// TIA Portal project "000_empty" (V21)

(* hardware
DEVICE "PLC_1"  S7-1500 station
   slot 0: "Rail_0"  Rack  6ES7 590-1***0-0AA0
   slot 1: "PLC_1"  CPU 1513-1 PN  6ES7 513-1AL02-0AB0  V2.9
      slot 3: "CPU display_1"  6ES7591-1AA00-0AA0
      slot 32768: "PROFINET interface_1"  X1
         slot 32769: "Port_1"  X1 P1
         slot 32770: "Port_2"  X1 P2
      slot 34817: "Virtual CP interface port_1"  Virtual CP interface port  Virtual CP interface port
DEVICE "HMI_TP900"  TP900 Comfort
   slot 0: "HMI_TP900"  TP900 Comfort  6AV2 124-0JC01-0AX0  17.0.0.0
   slot 1: "HMI_TP900"  TP900 Comfort  6AV2 124-0JC01-0AX0  17.0.0.0
   slot 5: "HMI_TP900.IE_CP_1"  PROFINET Interface  17.0.0.0
      slot 1: "PROFINET Interface_1"  PROFINET Interface
         slot 1: "Port_1"  Port
         slot 2: "Port_2"  Port
   slot 7: "HMI_TP900.MPI/DP_CP_1"  MPI/DP Interface  17.0.0.0
DEVICE "HMI_PCADV"  SIMATIC PC station
   slot 0: "SIMATIC PC station"  Rail  SIMATIC PC-Station  V1.0
      slot 125: "Stationmanager"  Station_Manager  V6.0.4
   slot 1: "HMI_RT_1"  WinCC RT Advanced  6AV2 104-0xxxx-xxxx  17.0.0.0
      slot 33792: "Computer interface"  Host interface
   slot 2: "IE_general_1"  IE General  IE_CP  V8.2.0
      slot 1: "PROFINET interface"  IEGeneral.Interface.8.2.0
DEVICE "HMI_TP900S"  TP900 Comfort
   slot 0: "HMI_TP900S"  TP900 Comfort  6AV2 124-0JC01-0AX0  17.0.0.0
   slot 1: "HMI_TP900S"  TP900 Comfort  6AV2 124-0JC01-0AX0  17.0.0.0
   slot 5: "HMI_TP900S.IE_CP_1"  PROFINET Interface  17.0.0.0
      slot 1: "PROFINET Interface_1"  PROFINET Interface
         slot 1: "Port_1"  Port
         slot 2: "Port_2"  Port
   slot 7: "HMI_TP900S.MPI/DP_CP_1"  MPI/DP Interface  17.0.0.0
DEVICE "HMI_TP1200"  TP1200 Comfort
   slot 0: "HMI_TP1200"  TP1200 Comfort  6AV2 124-0MC01-0AX0  17.0.0.0
   slot 1: "HMI_TP1200"  TP1200 Comfort  6AV2 124-0MC01-0AX0  17.0.0.0
   slot 5: "HMI_TP1200.IE_CP_1"  PROFINET Interface  17.0.0.0
      slot 1: "PROFINET Interface_1"  PROFINET Interface
         slot 1: "Port_1"  Port
         slot 2: "Port_2"  Port
   slot 7: "HMI_TP1200.MPI/DP_CP_1"  MPI/DP Interface  17.0.0.0
*)

// ===== PLC "PLC_1"  CPU 1513-1 PN =====

VAR_GLOBAL   // PLC tag table "Default tag table"
   "Plc_Bool" AT %M100.0 : Bool;
   "Plc_Int" AT %MW102 : Int;
   "Plc_Real" AT %MD104 : Real;
   "Plc_Byte" AT %MB108 : Byte;
END_VAR

ORGANIZATION_BLOCK "Main"   // OB1, LAD, ProgramCycle
TITLE = "Main Program Sweep (Cycle)"
{ S7_Optimized_Access := 'TRUE' }
VERSION : 0.1
   VAR_INPUT
      Initial_Call : Bool;   // Initial call of this OB
      Remanence : Bool;   // =True, if remanent data are available
   END_VAR
BEGIN
END_ORGANIZATION_BLOCK

(* ===== HMI "HMI_TP900" =====
system functions are stored by id; their names below are inferred from use
connection "HMI_Connection_1": ETHERNET, S7_1500_OMS

HMI tags "Default tag table"
   "Hmi_Bool" : Bool, internal
   "Hmi_Int" : Int, internal
   "Hmi_Real" : Real, internal
   "Hmi_String" : WString[254], internal
   "Ext_Bool" : Bool = PLC Plc_Bool AT %M100.0, 1 s
   "Ext_Int" : Int = PLC Plc_Int AT %MW102, 1 s
   "Ext_Real" : Real = PLC Plc_Real AT %MD104, 1 s
   "Ext_Byte" : Byte = PLC Plc_Byte AT %MB108, 1 s

HMI tags "C03_Tags"
   "D_State" : Int, internal
   "D_Bool" : Bool, internal
   "D_SInt" : SInt, internal
   "D_Int" : Int, internal
   "D_DInt" : DInt, internal
   "D_USInt" : USInt, internal
   "D_UInt" : UInt, internal
   "D_UDInt" : UDInt, internal
   "D_Real" : Real, internal
   "D_LReal" : LReal, internal
   "D_String" : WString[254], internal
   "D_DateTime" : DateTime, internal
   "D_Pct" : Int, internal
   "D_Range" : Int, internal
   "D_Bits" : Int, internal
   "D_Vis" : Bool, internal
   "D_En" : Bool, internal
   "D_X" : Int, internal
   "D_Y" : Int, internal
   "D_Max" : Real, internal
   "D_Min" : Real, internal
   "D_TL" : Int, internal
   "D_BarR" : Real, internal

text list "TL_Value": -100..-1 'Negative (-100..-1)'; 0 'Zero'; 1..9 'One to nine'; 10 'Ten: Ünïcödé äöüß ÄÖÜ €'; 32000 'Undefined value (default entry)'

text list "TL_Bit": 0 'Off (0)'; 1 'On (1)'

text list "TL_BitNo": 0 'Bit 0 set'; 1 'Bit 1 set'; 2 'Bit 2 set'; 3 'Bit 3 set'

graphic list "GL_Bit": 0 'G_EMF'; 1 'G_WMF'

graphic list "GL_BitNo": 0 'G_PNG'; 1 'G_JPG'; 2 'G_BMP'; 3 'G_TIF'

graphic list "GL_Value": -100..-1 'G_GIF'; 0 'G_PNG'; 1..9 'G_JPG'; 10 'G_BMP'; 32000 'G_SVG'

SlideinScreen "GraphX_Slidein_Top" 800x120
   TextField "SI_Title" at 10,10 size 300x20; Text 'Slide-in screen Top'
   Bar "SI_Bar" at 330,10 size 200x40
      ProcessValue <- "D_Pct"
   IOField "SI_Value" at 560,10 size 120x30; FormatPattern s99999
      ProcessValue <- "D_Int"

screen "All_Objects" 800x480
   TextField "TextField_1" at 680,10 size 100x30; Text 'Text'
   GraphicView "GraphicView_1" at 10,80 size 100x60
   IOField "IOField_1" at 130,80 size 100x30
   Button "Button_1" at 250,80 size 100x40; TextOff 'Text'
   SymbolicIOField "SymbolicIOField_1" at 370,80 size 120x30; TextOff '0'; TextOn '1'
   GraphicIOField "GraphicIOField_1" at 510,80 size 60x60
   DateTimeField "DateTimeField_1" at 590,80 size 160x30
   Bar "Bar_1" at 10,160 size 40x120
   Switch "Switch_1" at 70,160 size 120x40; CaptionText 'Switch'; TextOff '0'; TextOn '1'
   SymbolLibrary "SymbolLibrary_1" at 210,160 size 60x60
   Slider "Slider_1" at 290,160 size 60x160; Caption 'SIMATIC'
   Gauge "Gauge_1" at 370,160 size 150x150; CaptionText 'SIMATIC'
   Clock "Clock_1" at 540,160 size 150x150

screen "Ctl_01_AlarmView" 800x480, template "Nav"
   AlarmView "Alarm view_1" at 3,3 size 600x300

screen "Ctl_02_TrendView" 800x480, template "Nav"
   TrendView "Trend view_1" at 3,3 size 600x300

screen "Ctl_03_UserView" 800x480, template "Nav"
   UserView "User view_1" at 3,3 size 480x240

screen "Ctl_04_HtmlBrowser" 800x480, template "Nav"
   HTMLBrowser "HTML browser_1" at 3,3 size 192x192

screen "Ctl_05_WatchTable" 800x480, template "Nav"
   StatusForce "Watch table_1" at 3,3 size 600x300; ToolTipText 'Text'

screen "Ctl_06_SmartClientView" 800x480, template "Nav"
   SmartClientView "Sm@rtClient view_1" at 3,3 size 320x240

screen "Ctl_07_RecipeView" 800x480, template "Nav"
   RecipeView "Recipe view_1" at 3,3 size 400x330

screen "Ctl_09_SysDiagView" 800x480, template "Nav"
   SysDiagControl "System diagnostics view_1" at 3,3 size 600x300

screen "Ctl_10_MediaPlayer" 800x480, template "Nav"
   MediaPlayer "Media Player_1" at 3,3 size 240x240

screen "Ctl_15_CameraView" 800x480, template "Nav"
   CameraControl "Camera view_1" at 3,3 size 320x240

screen "Ctl_16_PdfView" 800x480, template "Nav"
   PDFView "PDFView_1" at 3,3 size 320x240

Template "Nav" 800x480
   Button "Nav_01" at 770,2 size 28x22; TextOff 'Text'
      on Click: ActivateScreen("Ctl_01_AlarmView", 0)
   Button "Nav_02" at 770,28 size 28x22; TextOff 'Text'
      on Click: ActivateScreen("Ctl_02_TrendView", 0)
   Button "Nav_03" at 770,54 size 28x22; TextOff 'Text'
      on Click: ActivateScreen("Ctl_03_UserView", 0)
   Button "Nav_04" at 770,80 size 28x22; TextOff 'Text'
      on Click: ActivateScreen("Ctl_04_HtmlBrowser", 0)
   Button "Nav_05" at 770,106 size 28x22; TextOff 'Text'
      on Click: ActivateScreen("Ctl_05_WatchTable", 0)
   Button "Nav_06" at 770,132 size 28x22; TextOff 'Text'
      on Click: ActivateScreen("Ctl_06_SmartClientView", 0)
   Button "Nav_07" at 770,158 size 28x22; TextOff 'Text'
      on Click: ActivateScreen("Ctl_07_RecipeView", 0)
   Button "Nav_09" at 770,210 size 28x22; TextOff 'Text'
      on Click: ActivateScreen("Ctl_09_SysDiagView", 0)
   Button "Nav_10" at 770,236 size 28x22; TextOff 'Text'
      on Click: ActivateScreen("Ctl_10_MediaPlayer", 0)
   Button "Nav_15" at 770,366 size 28x22; TextOff 'Text'
      on Click: ActivateScreen("Ctl_15_CameraView", 0)
   Button "Nav_16" at 770,392 size 28x22; TextOff 'Text'
      on Click: ActivateScreen("Ctl_16_PdfView", 0)
   Button "Nav_17" at 770,418 size 28x22; TextOff 'Text'
      on Click: ActivateScreen("All_Objects", 0)

screen "P_Line_1" 800x480
   TextField "Label_Default" at 10,62 size 108x16; Text 'Default'
   TextField "Label_BackColor" at 120,62 size 108x16; Text 'BackColor'
   TextField "Label_Color" at 230,62 size 108x16; Text 'Color'
   TextField "Label_EndStyle" at 340,62 size 108x16; Text 'EndStyle'
   TextField "Label_EndStyle_2" at 450,62 size 108x16; Text 'EndStyle_2'
   TextField "Label_EndStyle_3" at 560,62 size 108x16; Text 'EndStyle_3'
   TextField "Label_EndStyle_4" at 670,62 size 108x16; Text 'EndStyle_4'
   TextField "Label_EndStyle_5" at 10,138 size 108x16; Text 'EndStyle_5'
   TextField "Label_FillStyle" at 120,138 size 108x16; Text 'FillStyle'
   TextField "Label_Flashing" at 230,138 size 108x16; Text 'Flashing'
   TextField "Label_LineEndShapeStyle_2" at 340,138 size 108x16; Text 'LineEndShapeStyle_2'
   TextField "Label_LineWidth" at 450,138 size 108x16; Text 'LineWidth'
   TextField "Label_StartStyle" at 560,138 size 108x16; Text 'StartStyle'
   TextField "Label_StartStyle_2" at 670,138 size 108x16; Text 'StartStyle_2'
   TextField "Label_StartStyle_3" at 10,214 size 108x16; Text 'StartStyle_3'
   TextField "Label_StartStyle_4" at 120,214 size 108x16; Text 'StartStyle_4'
   TextField "Label_StartStyle_5" at 230,214 size 108x16; Text 'StartStyle_5'
   TextField "Label_Style" at 340,214 size 108x16; Text 'Style'
   TextField "Label_Style_2" at 450,214 size 108x16; Text 'Style_2'
   TextField "Label_Style_3" at 560,214 size 108x16; Text 'Style_3'
   TextField "Label_Style_4" at 670,214 size 108x16; Text 'Style_4'
   TextField "Label_UseDesignColorSchema" at 10,290 size 108x16; Text 'UseDesignColorSchema'
   Button "Next" at 758,456 size 40x22; TextOff 'Text'
      on Click: ActivateScreen("P_Polyline_1", 0)

screen "P_Polyline_1" 800x480
   TextField "Label_Default" at 10,62 size 108x16; Text 'Default'
   TextField "Label_BackColor" at 120,62 size 108x16; Text 'BackColor'
   TextField "Label_Color" at 230,62 size 108x16; Text 'Color'
   TextField "Label_EndStyle" at 340,62 size 108x16; Text 'EndStyle'
   TextField "Label_EndStyle_2" at 450,62 size 108x16; Text 'EndStyle_2'
   TextField "Label_EndStyle_3" at 560,62 size 108x16; Text 'EndStyle_3'
   TextField "Label_EndStyle_4" at 670,62 size 108x16; Text 'EndStyle_4'
   TextField "Label_EndStyle_5" at 10,138 size 108x16; Text 'EndStyle_5'
   TextField "Label_FillStyle" at 120,138 size 108x16; Text 'FillStyle'
   TextField "Label_Flashing" at 230,138 size 108x16; Text 'Flashing'
   TextField "Label_LineEndShapeStyle_2" at 340,138 size 108x16; Text 'LineEndShapeStyle_2'
   TextField "Label_LineWidth" at 450,138 size 108x16; Text 'LineWidth'
   TextField "Label_StartStyle" at 560,138 size 108x16; Text 'StartStyle'
   TextField "Label_StartStyle_2" at 670,138 size 108x16; Text 'StartStyle_2'
   TextField "Label_StartStyle_3" at 10,214 size 108x16; Text 'StartStyle_3'
   TextField "Label_StartStyle_4" at 120,214 size 108x16; Text 'StartStyle_4'
   TextField "Label_StartStyle_5" at 230,214 size 108x16; Text 'StartStyle_5'
   TextField "Label_Style" at 340,214 size 108x16; Text 'Style'
   TextField "Label_Style_2" at 450,214 size 108x16; Text 'Style_2'
   TextField "Label_Style_3" at 560,214 size 108x16; Text 'Style_3'
   TextField "Label_Style_4" at 670,214 size 108x16; Text 'Style_4'
   TextField "Label_UseDesignColorSchema" at 10,290 size 108x16; Text 'UseDesignColorSchema'
   Button "Next" at 758,456 size 40x22; TextOff 'Text'
      on Click: ActivateScreen("P_Polygon_1", 0)

screen "P_Polygon_1" 800x480
   TextField "Label_Default" at 10,62 size 108x16; Text 'Default'
   TextField "Label_BackColor" at 120,62 size 108x16; Text 'BackColor'
   TextField "Label_BackFillStyle" at 230,62 size 108x16; Text 'BackFillStyle'
   TextField "Label_BorderColor" at 340,62 size 108x16; Text 'BorderColor'
   TextField "Label_BorderWidth" at 450,62 size 108x16; Text 'BorderWidth'
   TextField "Label_EdgeStyle" at 560,62 size 108x16; Text 'EdgeStyle'
   TextField "Label_EdgeStyle_2" at 670,62 size 108x16; Text 'EdgeStyle_2'
   TextField "Label_EdgeStyle_3" at 10,138 size 108x16; Text 'EdgeStyle_3'
   TextField "Label_EdgeStyle_4" at 120,138 size 108x16; Text 'EdgeStyle_4'
   TextField "Label_Flashing" at 230,138 size 108x16; Text 'Flashing'
   TextField "Label_UseDesignColorSchema" at 340,138 size 108x16; Text 'UseDesignColorSchema'
   Button "Next" at 758,456 size 40x22; TextOff 'Text'
      on Click: ActivateScreen("P_Ellipse_1", 0)

screen "P_Ellipse_1" 800x480
   TextField "Label_Default" at 10,62 size 108x16; Text 'Default'
   TextField "Label_BackColor" at 120,62 size 108x16; Text 'BackColor'
   TextField "Label_BackFillStyle" at 230,62 size 108x16; Text 'BackFillStyle'
   TextField "Label_BorderColor" at 340,62 size 108x16; Text 'BorderColor'
   TextField "Label_BorderWidth" at 450,62 size 108x16; Text 'BorderWidth'
   TextField "Label_EdgeStyle" at 560,62 size 108x16; Text 'EdgeStyle'
   TextField "Label_EdgeStyle_2" at 670,62 size 108x16; Text 'EdgeStyle_2'
   TextField "Label_EdgeStyle_3" at 10,138 size 108x16; Text 'EdgeStyle_3'
   TextField "Label_EdgeStyle_4" at 120,138 size 108x16; Text 'EdgeStyle_4'
   TextField "Label_Flashing" at 230,138 size 108x16; Text 'Flashing'
   TextField "Label_UseDesignColorSchema" at 340,138 size 108x16; Text 'UseDesignColorSchema'
   Button "Next" at 758,456 size 40x22; TextOff 'Text'
      on Click: ActivateScreen("P_Circle_1", 0)

screen "P_Circle_1" 800x480
   TextField "Label_Default" at 10,62 size 58x16; Text 'Default'
   TextField "Label_BackColor" at 70,62 size 58x16; Text 'BackColor'
   TextField "Label_BackFillStyle" at 130,62 size 58x16; Text 'BackFillStyle'
   TextField "Label_BorderColor" at 190,62 size 58x16; Text 'BorderColor'
   TextField "Label_BorderWidth" at 250,62 size 58x16; Text 'BorderWidth'
   TextField "Label_EdgeStyle" at 310,62 size 58x16; Text 'EdgeStyle'
   TextField "Label_EdgeStyle_2" at 370,62 size 58x16; Text 'EdgeStyle_2'
   TextField "Label_EdgeStyle_3" at 430,62 size 58x16; Text 'EdgeStyle_3'
   TextField "Label_EdgeStyle_4" at 490,62 size 58x16; Text 'EdgeStyle_4'
   TextField "Label_Flashing" at 550,62 size 58x16; Text 'Flashing'
   TextField "Label_UseDesignColorSchema" at 610,62 size 58x16; Text 'UseDesignColorSchema'
   Button "Next" at 758,456 size 40x22; TextOff 'Text'
      on Click: ActivateScreen("P_Rectangle_1", 0)

screen "P_Rectangle_1" 800x480
   TextField "Label_Default" at 10,62 size 108x16; Text 'Default'
   TextField "Label_BackColor" at 120,62 size 108x16; Text 'BackColor'
   TextField "Label_BackFillStyle" at 230,62 size 108x16; Text 'BackFillStyle'
   TextField "Label_BorderColor" at 340,62 size 108x16; Text 'BorderColor'
   TextField "Label_BorderWidth" at 450,62 size 108x16; Text 'BorderWidth'
   TextField "Label_EdgeStyle" at 560,62 size 108x16; Text 'EdgeStyle'
   TextField "Label_EdgeStyle_2" at 670,62 size 108x16; Text 'EdgeStyle_2'
   TextField "Label_EdgeStyle_3" at 10,138 size 108x16; Text 'EdgeStyle_3'
   TextField "Label_EdgeStyle_4" at 120,138 size 108x16; Text 'EdgeStyle_4'
   TextField "Label_Flashing" at 230,138 size 108x16; Text 'Flashing'
   TextField "Label_RoundCornerHeight" at 340,138 size 108x16; Text 'RoundCornerHeight'
   TextField "Label_RoundCornerWidth" at 450,138 size 108x16; Text 'RoundCornerWidth'
   TextField "Label_UseDesignColorSchema" at 560,138 size 108x16; Text 'UseDesignColorSchema'
   Button "Next" at 758,456 size 40x22; TextOff 'Text'
      on Click: ActivateScreen("P_TextField_1", 0)

screen "P_TextField_1" 800x480
   TextField "Default" at 10,10 size 100x30; Text 'Text'
   TextField "Label_Default" at 10,42 size 108x16; Text 'Default'
   TextField "BackColor" at 120,10 size 100x30; Text 'Text'
   TextField "Label_BackColor" at 120,42 size 108x16; Text 'BackColor'
   TextField "BackFillStyle" at 230,10 size 100x30; Text 'Text'
   TextField "Label_BackFillStyle" at 230,42 size 108x16; Text 'BackFillStyle'
   TextField "BorderBackColor" at 340,10 size 100x30; Text 'Text'
   TextField "Label_BorderBackColor" at 340,42 size 108x16; Text 'BorderBackColor'
   TextField "BorderColor" at 450,10 size 100x30; Text 'Text'
   TextField "Label_BorderColor" at 450,42 size 108x16; Text 'BorderColor'
   TextField "BorderWidth" at 560,10 size 100x30; Text 'Text'
   TextField "Label_BorderWidth" at 560,42 size 108x16; Text 'BorderWidth'
   TextField "BottomMargin" at 670,10 size 100x30; Text 'Text'
   TextField "Label_BottomMargin" at 670,42 size 108x16; Text 'BottomMargin'
   TextField "CornerRadius" at 10,66 size 100x30; Text 'Text'
   TextField "Label_CornerRadius" at 10,98 size 108x16; Text 'CornerRadius'
   TextField "EdgeStyle" at 120,66 size 100x30; Text 'Text'
   TextField "Label_EdgeStyle" at 120,98 size 108x16; Text 'EdgeStyle'
   TextField "EdgeStyle_2" at 230,66 size 100x30; Text 'Text'
   TextField "Label_EdgeStyle_2" at 230,98 size 108x16; Text 'EdgeStyle_2'
   TextField "EdgeStyle_3" at 340,66 size 100x30; Text 'Text'
   TextField "Label_EdgeStyle_3" at 340,98 size 108x16; Text 'EdgeStyle_3'
   TextField "EdgeStyle_4" at 450,66 size 100x30; Text 'Text'
   TextField "Label_EdgeStyle_4" at 450,98 size 108x16; Text 'EdgeStyle_4'
   TextField "FitToLargest" at 560,66 size 100x30; Text 'Text'
   TextField "Label_FitToLargest" at 560,98 size 108x16; Text 'FitToLargest'
   TextField "Flashing" at 670,66 size 100x30; Text 'Text'
   TextField "Label_Flashing" at 670,98 size 108x16; Text 'Flashing'
   TextField "ForeColor" at 10,122 size 100x30; Text 'Text'
   TextField "Label_ForeColor" at 10,154 size 108x16; Text 'ForeColor'
   TextField "HorizontalAlignment" at 120,122 size 100x30; Text 'Text'
   TextField "Label_HorizontalAlignment" at 120,154 size 108x16; Text 'HorizontalAlignment'
   TextField "HorizontalAlignment_2" at 230,122 size 100x30; Text 'Text'
   TextField "Label_HorizontalAlignment_2" at 230,154 size 108x16; Text 'HorizontalAlignment_2'
   TextField "LeftMargin" at 340,122 size 100x30; Text 'Text'
   TextField "Label_LeftMargin" at 340,154 size 108x16; Text 'LeftMargin'
   TextField "RightMargin" at 450,122 size 100x30; Text 'Text'
   TextField "Label_RightMargin" at 450,154 size 108x16; Text 'RightMargin'
   TextField "TopMargin" at 560,122 size 100x30; Text 'Text'
   TextField "Label_TopMargin" at 560,154 size 108x16; Text 'TopMargin'
   TextField "UseDesignColorSchema" at 670,122 size 100x30; Text 'Text'
   TextField "Label_UseDesignColorSchema" at 670,154 size 108x16; Text 'UseDesignColorSchema'
   TextField "VerticalAlignment" at 10,178 size 100x30; Text 'Text'
   TextField "Label_VerticalAlignment" at 10,210 size 108x16; Text 'VerticalAlignment'
   TextField "VerticalAlignment_2" at 120,178 size 100x30; Text 'Text'
   TextField "Label_VerticalAlignment_2" at 120,210 size 108x16; Text 'VerticalAlignment_2'
   Button "Next" at 758,456 size 40x22; TextOff 'Text'
      on Click: ActivateScreen("P_GraphicView_1", 0)

screen "P_GraphicView_1" 800x480
   GraphicView "Default" at 10,10 size 100x60
   TextField "Label_Default" at 10,72 size 108x16; Text 'Default'
   GraphicView "BackColor" at 120,10 size 100x60
   TextField "Label_BackColor" at 120,72 size 108x16; Text 'BackColor'
   GraphicView "BackFillStyle" at 230,10 size 100x60
   TextField "Label_BackFillStyle" at 230,72 size 108x16; Text 'BackFillStyle'
   GraphicView "BorderColor" at 340,10 size 100x60
   TextField "Label_BorderColor" at 340,72 size 108x16; Text 'BorderColor'
   GraphicView "BorderWidth" at 450,10 size 100x60
   TextField "Label_BorderWidth" at 450,72 size 108x16; Text 'BorderWidth'
   GraphicView "EdgeStyle" at 560,10 size 100x60
   TextField "Label_EdgeStyle" at 560,72 size 108x16; Text 'EdgeStyle'
   GraphicView "EdgeStyle_2" at 670,10 size 100x60
   TextField "Label_EdgeStyle_2" at 670,72 size 108x16; Text 'EdgeStyle_2'
   GraphicView "EdgeStyle_3" at 10,96 size 100x60
   TextField "Label_EdgeStyle_3" at 10,158 size 108x16; Text 'EdgeStyle_3'
   GraphicView "EdgeStyle_4" at 120,96 size 100x60
   TextField "Label_EdgeStyle_4" at 120,158 size 108x16; Text 'EdgeStyle_4'
   GraphicView "FitToLargest" at 230,96 size 100x60
   TextField "Label_FitToLargest" at 230,158 size 108x16; Text 'FitToLargest'
   GraphicView "Flashing" at 340,96 size 100x60
   TextField "Label_Flashing" at 340,158 size 108x16; Text 'Flashing'
   GraphicView "TransparentColor" at 450,96 size 100x60
   TextField "Label_TransparentColor" at 450,158 size 108x16; Text 'TransparentColor'
   GraphicView "UseTransparentColor" at 560,96 size 100x60
   TextField "Label_UseTransparentColor" at 560,158 size 108x16; Text 'UseTransparentColor'
   Button "Next" at 758,456 size 40x22; TextOff 'Text'
      on Click: ActivateScreen("P_IOField_1", 0)

screen "P_Button_1" 800x480
   Button "Default" at 10,10 size 100x40; TextOff 'Text'
   TextField "Label_Default" at 10,52 size 108x16; Text 'Default'
   Button "BackColor" at 120,10 size 100x40; TextOff 'Text'
   TextField "Label_BackColor" at 120,52 size 108x16; Text 'BackColor'
   Button "BackFillStyle" at 230,10 size 100x40; TextOff 'Text'
   TextField "Label_BackFillStyle" at 230,52 size 108x16; Text 'BackFillStyle'
   Button "BorderBackColor" at 340,10 size 100x40; TextOff 'Text'
   TextField "Label_BorderBackColor" at 340,52 size 108x16; Text 'BorderBackColor'
   Button "BorderColor" at 450,10 size 100x40; TextOff 'Text'
   TextField "Label_BorderColor" at 450,52 size 108x16; Text 'BorderColor'
   Button "BorderWidth" at 560,10 size 100x40; TextOff 'Text'
   TextField "Label_BorderWidth" at 560,52 size 108x16; Text 'BorderWidth'
   Button "CornerRadius" at 670,10 size 100x40; TextOff 'Text'
   TextField "Label_CornerRadius" at 670,52 size 108x16; Text 'CornerRadius'
   Button "EdgeStyle" at 10,76 size 100x40; TextOff 'Text'
   TextField "Label_EdgeStyle" at 10,118 size 108x16; Text 'EdgeStyle'
   Button "EdgeStyle_2" at 120,76 size 100x40; TextOff 'Text'
   TextField "Label_EdgeStyle_2" at 120,118 size 108x16; Text 'EdgeStyle_2'
   Button "EdgeStyle_3" at 230,76 size 100x40; TextOff 'Text'
   TextField "Label_EdgeStyle_3" at 230,118 size 108x16; Text 'EdgeStyle_3'
   Button "EdgeStyle_4" at 340,76 size 100x40; TextOff 'Text'
   TextField "Label_EdgeStyle_4" at 340,118 size 108x16; Text 'EdgeStyle_4'
   Button "FirstGradientColor" at 450,76 size 100x40; TextOff 'Text'
   TextField "Label_FirstGradientColor" at 450,118 size 108x16; Text 'FirstGradientColor'
   Button "FirstGradientOffset" at 560,76 size 100x40; TextOff 'Text'
   TextField "Label_FirstGradientOffset" at 560,118 size 108x16; Text 'FirstGradientOffset'
   Button "FitToLargest" at 670,76 size 100x40; TextOff 'Text'
   TextField "Label_FitToLargest" at 670,118 size 108x16; Text 'FitToLargest'
   Button "Flashing" at 10,142 size 100x40; TextOff 'Text'
   TextField "Label_Flashing" at 10,184 size 108x16; Text 'Flashing'
   Button "FocusColor" at 120,142 size 100x40; TextOff 'Text'
   TextField "Label_FocusColor" at 120,184 size 108x16; Text 'FocusColor'
   Button "FocusWidth" at 230,142 size 100x40; TextOff 'Text'
   TextField "Label_FocusWidth" at 230,184 size 108x16; Text 'FocusWidth'
   Button "ForeColor" at 340,142 size 100x40; TextOff 'Text'
   TextField "Label_ForeColor" at 340,184 size 108x16; Text 'ForeColor'
   Button "HorizontalAlignment" at 450,142 size 100x40; TextOff 'Text'
   TextField "Label_HorizontalAlignment" at 450,184 size 108x16; Text 'HorizontalAlignment'
   Button "HorizontalAlignment_2" at 560,142 size 100x40; TextOff 'Text'
   TextField "Label_HorizontalAlignment_2" at 560,184 size 108x16; Text 'HorizontalAlignment_2'
   Button "HorizontalPictureAlignment" at 670,142 size 100x40; TextOff 'Text'
   TextField "Label_HorizontalPictureAlignment" at 670,184 size 108x16; Text 'HorizontalPictureAlignment'
   Button "HorizontalPictureAlignment_2" at 10,208 size 100x40; TextOff 'Text'
   TextField "Label_HorizontalPictureAlignment_2" at 10,250 size 108x16; Text 'HorizontalPictureAlignment_2'
   Button "MiddleGradientColor" at 120,208 size 100x40; TextOff 'Text'
   TextField "Label_MiddleGradientColor" at 120,250 size 108x16; Text 'MiddleGradientColor'
   Button "Mode_5" at 230,208 size 100x40; TextOff 'Text'
   TextField "Label_Mode_5" at 230,250 size 108x16; Text 'Mode_5'
   Button "Mode_7" at 340,208 size 100x40; TextOff 'Text'
   TextField "Label_Mode_7" at 340,250 size 108x16; Text 'Mode_7'
   Button "PictureAreaBottomMargin" at 450,208 size 100x40; TextOff 'Text'
   TextField "Label_PictureAreaBottomMargin" at 450,250 size 108x16; Text 'PictureAreaBottomMargin'
   Button "PictureAreaLeftMargin" at 560,208 size 100x40; TextOff 'Text'
   TextField "Label_PictureAreaLeftMargin" at 560,250 size 108x16; Text 'PictureAreaLeftMargin'
   Button "PictureAreaRightMargin" at 670,208 size 100x40; TextOff 'Text'
   TextField "Label_PictureAreaRightMargin" at 670,250 size 108x16; Text 'PictureAreaRightMargin'
   Button "PictureAreaTopMargin" at 10,274 size 100x40; TextOff 'Text'
   TextField "Label_PictureAreaTopMargin" at 10,316 size 108x16; Text 'PictureAreaTopMargin'
   Button "SecondGradientColor" at 120,274 size 100x40; TextOff 'Text'
   TextField "Label_SecondGradientColor" at 120,316 size 108x16; Text 'SecondGradientColor'
   Button "SecondGradientOffset" at 230,274 size 100x40; TextOff 'Text'
   TextField "Label_SecondGradientOffset" at 230,316 size 108x16; Text 'SecondGradientOffset'
   Button "TextAreaBottomMargin" at 340,274 size 100x40; TextOff 'Text'
   TextField "Label_TextAreaBottomMargin" at 340,316 size 108x16; Text 'TextAreaBottomMargin'
   Button "TextAreaLeftMargin" at 450,274 size 100x40; TextOff 'Text'
   TextField "Label_TextAreaLeftMargin" at 450,316 size 108x16; Text 'TextAreaLeftMargin'
   Button "TextAreaRightMargin" at 560,274 size 100x40; TextOff 'Text'
   TextField "Label_TextAreaRightMargin" at 560,316 size 108x16; Text 'TextAreaRightMargin'
   Button "TextAreaTopMargin" at 670,274 size 100x40; TextOff 'Text'
   TextField "Label_TextAreaTopMargin" at 670,316 size 108x16; Text 'TextAreaTopMargin'
   Button "UseDesignColorSchema" at 10,340 size 100x40; TextOff 'Text'
   TextField "Label_UseDesignColorSchema" at 10,382 size 108x16; Text 'UseDesignColorSchema'
   Button "UseFirstGradient" at 120,340 size 100x40; TextOff 'Text'
   TextField "Label_UseFirstGradient" at 120,382 size 108x16; Text 'UseFirstGradient'
   Button "UseSecondGradient" at 230,340 size 100x40; TextOff 'Text'
   TextField "Label_UseSecondGradient" at 230,382 size 108x16; Text 'UseSecondGradient'
   Button "VerticalAlignment" at 340,340 size 100x40; TextOff 'Text'
   TextField "Label_VerticalAlignment" at 340,382 size 108x16; Text 'VerticalAlignment'
   Button "VerticalAlignment_2" at 450,340 size 100x40; TextOff 'Text'
   TextField "Label_VerticalAlignment_2" at 450,382 size 108x16; Text 'VerticalAlignment_2'
   Button "VerticalPictureAlignment" at 560,340 size 100x40; TextOff 'Text'
   TextField "Label_VerticalPictureAlignment" at 560,382 size 108x16; Text 'VerticalPictureAlignment'
   Button "VerticalPictureAlignment_2" at 670,340 size 100x40; TextOff 'Text'
   TextField "Label_VerticalPictureAlignment_2" at 670,382 size 108x16; Text 'VerticalPictureAlignment_2'
   Button "Next" at 758,456 size 40x22; TextOff 'Text'
      on Click: ActivateScreen("P_SymbolicIOField_1", 0)

screen "P_SymbolicIOField_1" 800x480
   SymbolicIOField "Default" at 10,10 size 120x30; TextOff '0'; TextOn '1'
   TextField "Label_Default" at 10,42 size 128x16; Text 'Default'
   SymbolicIOField "AboveUpperLimitColor" at 140,10 size 120x30; TextOff '0'; TextOn '1'
   TextField "Label_AboveUpperLimitColor" at 140,42 size 128x16; Text 'AboveUpperLimitColor'
   SymbolicIOField "BackColor" at 270,10 size 120x30; TextOff '0'; TextOn '1'
   TextField "Label_BackColor" at 270,42 size 128x16; Text 'BackColor'
   SymbolicIOField "BackFillStyle" at 400,10 size 120x30; TextOff '0'; TextOn '1'
   TextField "Label_BackFillStyle" at 400,42 size 128x16; Text 'BackFillStyle'
   SymbolicIOField "BelowLowerLimitColor" at 530,10 size 120x30; TextOff '0'; TextOn '1'
   TextField "Label_BelowLowerLimitColor" at 530,42 size 128x16; Text 'BelowLowerLimitColor'
   SymbolicIOField "BorderBackColor" at 660,10 size 120x30; TextOff '0'; TextOn '1'
   TextField "Label_BorderBackColor" at 660,42 size 128x16; Text 'BorderBackColor'
   SymbolicIOField "BorderColor" at 10,66 size 120x30; TextOff '0'; TextOn '1'
   TextField "Label_BorderColor" at 10,98 size 128x16; Text 'BorderColor'
   SymbolicIOField "BorderWidth" at 140,66 size 120x30; TextOff '0'; TextOn '1'
   TextField "Label_BorderWidth" at 140,98 size 128x16; Text 'BorderWidth'
   SymbolicIOField "BottomMargin" at 270,66 size 120x30; TextOff '0'; TextOn '1'
   TextField "Label_BottomMargin" at 270,98 size 128x16; Text 'BottomMargin'
   SymbolicIOField "CornerRadius" at 400,66 size 120x30; TextOff '0'; TextOn '1'
   TextField "Label_CornerRadius" at 400,98 size 128x16; Text 'CornerRadius'
   SymbolicIOField "CountVisibleItems" at 530,66 size 120x30; TextOff '0'; TextOn '1'
   TextField "Label_CountVisibleItems" at 530,98 size 128x16; Text 'CountVisibleItems'
   SymbolicIOField "EdgeStyle" at 660,66 size 120x30; TextOff '0'; TextOn '1'
   TextField "Label_EdgeStyle" at 660,98 size 128x16; Text 'EdgeStyle'
   SymbolicIOField "EdgeStyle_2" at 10,122 size 120x30; TextOff '0'; TextOn '1'
   TextField "Label_EdgeStyle_2" at 10,154 size 128x16; Text 'EdgeStyle_2'
   SymbolicIOField "EdgeStyle_3" at 140,122 size 120x30; TextOff '0'; TextOn '1'
   TextField "Label_EdgeStyle_3" at 140,154 size 128x16; Text 'EdgeStyle_3'
   SymbolicIOField "EdgeStyle_4" at 270,122 size 120x30; TextOff '0'; TextOn '1'
   TextField "Label_EdgeStyle_4" at 270,154 size 128x16; Text 'EdgeStyle_4'
   SymbolicIOField "EvenRowBackColor" at 400,122 size 120x30; TextOff '0'; TextOn '1'
   TextField "Label_EvenRowBackColor" at 400,154 size 128x16; Text 'EvenRowBackColor'
   SymbolicIOField "FitToLargest" at 530,122 size 120x30; TextOff '0'; TextOn '1'
   TextField "Label_FitToLargest" at 530,154 size 128x16; Text 'FitToLargest'
   SymbolicIOField "Flashing" at 660,122 size 120x30; TextOff '0'; TextOn '1'
   TextField "Label_Flashing" at 660,154 size 128x16; Text 'Flashing'
   SymbolicIOField "FlashingOnLimitViolation" at 10,178 size 120x30; TextOff '0'; TextOn '1'
   TextField "Label_FlashingOnLimitViolation" at 10,210 size 128x16; Text 'FlashingOnLimitViolation'
   SymbolicIOField "ForeColor" at 140,178 size 120x30; TextOff '0'; TextOn '1'
   TextField "Label_ForeColor" at 140,210 size 128x16; Text 'ForeColor'
   SymbolicIOField "HorizontalAlignment" at 270,178 size 120x30; TextOff '0'; TextOn '1'
   TextField "Label_HorizontalAlignment" at 270,210 size 128x16; Text 'HorizontalAlignment'
   SymbolicIOField "HorizontalAlignment_2" at 400,178 size 120x30; TextOff '0'; TextOn '1'
   TextField "Label_HorizontalAlignment_2" at 400,210 size 128x16; Text 'HorizontalAlignment_2'
   SymbolicIOField "LeftMargin" at 530,178 size 120x30; TextOff '0'; TextOn '1'
   TextField "Label_LeftMargin" at 530,210 size 128x16; Text 'LeftMargin'
   SymbolicIOField "Mode" at 660,178 size 120x30; TextOff '0'; TextOn '1'
   TextField "Label_Mode" at 660,210 size 128x16; Text 'Mode'
   SymbolicIOField "Mode_2" at 10,234 size 120x30; TextOff '0'; TextOn '1'
   TextField "Label_Mode_2" at 10,266 size 128x16; Text 'Mode_2'
   SymbolicIOField "RightMargin" at 140,234 size 120x30; TextOff '0'; TextOn '1'
   TextField "Label_RightMargin" at 140,266 size 128x16; Text 'RightMargin'
   SymbolicIOField "SelectBackColor" at 270,234 size 120x30; TextOff '0'; TextOn '1'
   TextField "Label_SelectBackColor" at 270,266 size 128x16; Text 'SelectBackColor'
   SymbolicIOField "SelectForeColor" at 400,234 size 120x30; TextOff '0'; TextOn '1'
   TextField "Label_SelectForeColor" at 400,266 size 128x16; Text 'SelectForeColor'
   SymbolicIOField "ShowDropDownButton" at 530,234 size 120x30; TextOff '0'; TextOn '1'
   TextField "Label_ShowDropDownButton" at 530,266 size 128x16; Text 'ShowDropDownButton'
   SymbolicIOField "ShowDropDownList" at 660,234 size 120x30; TextOff '0'; TextOn '1'
   TextField "Label_ShowDropDownList" at 660,266 size 128x16; Text 'ShowDropDownList'
   SymbolicIOField "TopMargin" at 10,290 size 120x30; TextOff '0'; TextOn '1'
   TextField "Label_TopMargin" at 10,322 size 128x16; Text 'TopMargin'
   SymbolicIOField "UseDesignColorSchema" at 140,290 size 120x30; TextOff '0'; TextOn '1'
   TextField "Label_UseDesignColorSchema" at 140,322 size 128x16; Text 'UseDesignColorSchema'
   SymbolicIOField "VerticalAlignment" at 270,290 size 120x30; TextOff '0'; TextOn '1'
   TextField "Label_VerticalAlignment" at 270,322 size 128x16; Text 'VerticalAlignment'
   SymbolicIOField "VerticalAlignment_2" at 400,290 size 120x30; TextOff '0'; TextOn '1'
   TextField "Label_VerticalAlignment_2" at 400,322 size 128x16; Text 'VerticalAlignment_2'
   Button "Next" at 758,456 size 40x22; TextOff 'Text'
      on Click: ActivateScreen("P_GraphicIOField_1", 0)

screen "P_GraphicIOField_1" 800x480
   GraphicIOField "Default" at 10,10 size 60x60
   TextField "Label_Default" at 10,72 size 68x16; Text 'Default'
   GraphicIOField "AboveUpperLimitColor" at 80,10 size 60x60
   TextField "Label_AboveUpperLimitColor" at 80,72 size 68x16; Text 'AboveUpperLimitColor'
   GraphicIOField "BackColor" at 150,10 size 60x60
   TextField "Label_BackColor" at 150,72 size 68x16; Text 'BackColor'
   GraphicIOField "BackFillStyle" at 220,10 size 60x60
   TextField "Label_BackFillStyle" at 220,72 size 68x16; Text 'BackFillStyle'
   GraphicIOField "BelowLowerLimitColor" at 290,10 size 60x60
   TextField "Label_BelowLowerLimitColor" at 290,72 size 68x16; Text 'BelowLowerLimitColor'
   GraphicIOField "BorderColor" at 360,10 size 60x60
   TextField "Label_BorderColor" at 360,72 size 68x16; Text 'BorderColor'
   GraphicIOField "BorderWidth" at 430,10 size 60x60
   TextField "Label_BorderWidth" at 430,72 size 68x16; Text 'BorderWidth'
   GraphicIOField "EdgeStyle" at 500,10 size 60x60
   TextField "Label_EdgeStyle" at 500,72 size 68x16; Text 'EdgeStyle'
   GraphicIOField "EdgeStyle_2" at 570,10 size 60x60
   TextField "Label_EdgeStyle_2" at 570,72 size 68x16; Text 'EdgeStyle_2'
   GraphicIOField "EdgeStyle_3" at 640,10 size 60x60
   TextField "Label_EdgeStyle_3" at 640,72 size 68x16; Text 'EdgeStyle_3'
   GraphicIOField "EdgeStyle_4" at 710,10 size 60x60
   TextField "Label_EdgeStyle_4" at 710,72 size 68x16; Text 'EdgeStyle_4'
   GraphicIOField "FitToLargest" at 10,96 size 60x60
   TextField "Label_FitToLargest" at 10,158 size 68x16; Text 'FitToLargest'
   GraphicIOField "Flashing" at 80,96 size 60x60
   TextField "Label_Flashing" at 80,158 size 68x16; Text 'Flashing'
   GraphicIOField "FlashingOnLimitViolation" at 150,96 size 60x60
   TextField "Label_FlashingOnLimitViolation" at 150,158 size 68x16; Text 'FlashingOnLimitViolation'
   GraphicIOField "FocusColor" at 220,96 size 60x60
   TextField "Label_FocusColor" at 220,158 size 68x16; Text 'FocusColor'
   GraphicIOField "FocusWidth" at 290,96 size 60x60
   TextField "Label_FocusWidth" at 290,158 size 68x16; Text 'FocusWidth'
   GraphicIOField "Mode" at 360,96 size 60x60
   TextField "Label_Mode" at 360,158 size 68x16; Text 'Mode'
   GraphicIOField "Mode_2" at 430,96 size 60x60
   TextField "Label_Mode_2" at 430,158 size 68x16; Text 'Mode_2'
   GraphicIOField "ScrollBarOrientation" at 500,96 size 60x60
   TextField "Label_ScrollBarOrientation" at 500,158 size 68x16; Text 'ScrollBarOrientation'
   GraphicIOField "TransparentColor" at 570,96 size 60x60
   TextField "Label_TransparentColor" at 570,158 size 68x16; Text 'TransparentColor'
   GraphicIOField "UseTransparentColor" at 640,96 size 60x60
   TextField "Label_UseTransparentColor" at 640,158 size 68x16; Text 'UseTransparentColor'
   Button "Next" at 758,456 size 40x22; TextOff 'Text'
      on Click: ActivateScreen("P_DateTimeField_1", 0)

screen "P_DateTimeField_1" 800x480
   DateTimeField "Default" at 10,10 size 160x30
   TextField "Label_Default" at 10,42 size 168x16; Text 'Default'
   DateTimeField "BackColor" at 180,10 size 160x30
   TextField "Label_BackColor" at 180,42 size 168x16; Text 'BackColor'
   DateTimeField "BackFillStyle" at 350,10 size 160x30
   TextField "Label_BackFillStyle" at 350,42 size 168x16; Text 'BackFillStyle'
   DateTimeField "BorderBackColor" at 520,10 size 160x30
   TextField "Label_BorderBackColor" at 520,42 size 168x16; Text 'BorderBackColor'
   DateTimeField "BorderColor" at 10,66 size 160x30
   TextField "Label_BorderColor" at 10,98 size 168x16; Text 'BorderColor'
   DateTimeField "BorderWidth" at 180,66 size 160x30
   TextField "Label_BorderWidth" at 180,98 size 168x16; Text 'BorderWidth'
   DateTimeField "BottomMargin" at 350,66 size 160x30
   TextField "Label_BottomMargin" at 350,98 size 168x16; Text 'BottomMargin'
   DateTimeField "CornerRadius" at 520,66 size 160x30
   TextField "Label_CornerRadius" at 520,98 size 168x16; Text 'CornerRadius'
   DateTimeField "DisplaySystemTime" at 10,122 size 160x30
   TextField "Label_DisplaySystemTime" at 10,154 size 168x16; Text 'DisplaySystemTime'
   DateTimeField "EdgeStyle" at 180,122 size 160x30
   TextField "Label_EdgeStyle" at 180,154 size 168x16; Text 'EdgeStyle'
   DateTimeField "EdgeStyle_2" at 350,122 size 160x30
   TextField "Label_EdgeStyle_2" at 350,154 size 168x16; Text 'EdgeStyle_2'
   DateTimeField "EdgeStyle_3" at 520,122 size 160x30
   TextField "Label_EdgeStyle_3" at 520,154 size 168x16; Text 'EdgeStyle_3'
   DateTimeField "EdgeStyle_4" at 10,178 size 160x30
   TextField "Label_EdgeStyle_4" at 10,210 size 168x16; Text 'EdgeStyle_4'
   DateTimeField "FitToLargest" at 180,178 size 160x30
   TextField "Label_FitToLargest" at 180,210 size 168x16; Text 'FitToLargest'
   DateTimeField "Flashing" at 350,178 size 160x30
   TextField "Label_Flashing" at 350,210 size 168x16; Text 'Flashing'
   DateTimeField "ForeColor" at 520,178 size 160x30
   TextField "Label_ForeColor" at 520,210 size 168x16; Text 'ForeColor'
   DateTimeField "HorizontalAlignment" at 10,234 size 160x30
   TextField "Label_HorizontalAlignment" at 10,266 size 168x16; Text 'HorizontalAlignment'
   DateTimeField "HorizontalAlignment_2" at 180,234 size 160x30
   TextField "Label_HorizontalAlignment_2" at 180,266 size 168x16; Text 'HorizontalAlignment_2'
   DateTimeField "LeftMargin" at 350,234 size 160x30
   TextField "Label_LeftMargin" at 350,266 size 168x16; Text 'LeftMargin'
   DateTimeField "LongDateTimeFormat" at 520,234 size 160x30
   TextField "Label_LongDateTimeFormat" at 520,266 size 168x16; Text 'LongDateTimeFormat'
   DateTimeField "Mode_3" at 10,290 size 160x30
   TextField "Label_Mode_3" at 10,322 size 168x16; Text 'Mode_3'
   DateTimeField "RightMargin" at 180,290 size 160x30
   TextField "Label_RightMargin" at 180,322 size 168x16; Text 'RightMargin'
   DateTimeField "ShowDate" at 350,290 size 160x30
   TextField "Label_ShowDate" at 350,322 size 168x16; Text 'ShowDate'
   DateTimeField "ShowTime" at 520,290 size 160x30
   TextField "Label_ShowTime" at 520,322 size 168x16; Text 'ShowTime'
   DateTimeField "TopMargin" at 10,346 size 160x30
   TextField "Label_TopMargin" at 10,378 size 168x16; Text 'TopMargin'
   DateTimeField "UseDesignColorSchema" at 180,346 size 160x30
   TextField "Label_UseDesignColorSchema" at 180,378 size 168x16; Text 'UseDesignColorSchema'
   DateTimeField "VerticalAlignment" at 350,346 size 160x30
   TextField "Label_VerticalAlignment" at 350,378 size 168x16; Text 'VerticalAlignment'
   DateTimeField "VerticalAlignment_2" at 520,346 size 160x30
   TextField "Label_VerticalAlignment_2" at 520,378 size 168x16; Text 'VerticalAlignment_2'
   Button "Next" at 758,456 size 40x22; TextOff 'Text'
      on Click: ActivateScreen("P_Bar_1", 0)

screen "P_Bar_1" 800x480
   Bar "Default" at 10,10 size 40x120
   TextField "Label_Default" at 10,132 size 48x16; Text 'Default'
   Bar "BackColor" at 60,10 size 40x120
   TextField "Label_BackColor" at 60,132 size 48x16; Text 'BackColor'
   Bar "BarBackColor" at 110,10 size 40x120
   TextField "Label_BarBackColor" at 110,132 size 48x16; Text 'BarBackColor'
   Bar "BarEdgeStyle" at 160,10 size 40x120
   TextField "Label_BarEdgeStyle" at 160,132 size 48x16; Text 'BarEdgeStyle'
   Bar "BarEdgeStyle_2" at 210,10 size 40x120
   TextField "Label_BarEdgeStyle_2" at 210,132 size 48x16; Text 'BarEdgeStyle_2'
   Bar "BarOrientation" at 260,10 size 40x120
   TextField "Label_BarOrientation" at 260,132 size 48x16; Text 'BarOrientation'
   Bar "BarOrientation_2" at 310,10 size 40x120
   TextField "Label_BarOrientation_2" at 310,132 size 48x16; Text 'BarOrientation_2'
   Bar "BarOrientation_3" at 360,10 size 40x120
   TextField "Label_BarOrientation_3" at 360,132 size 48x16; Text 'BarOrientation_3'
   Bar "BorderBackColor" at 410,10 size 40x120
   TextField "Label_BorderBackColor" at 410,132 size 48x16; Text 'BorderBackColor'
   Bar "BorderColor" at 460,10 size 40x120
   TextField "Label_BorderColor" at 460,132 size 48x16; Text 'BorderColor'
   Bar "BorderWidth" at 510,10 size 40x120
   TextField "Label_BorderWidth" at 510,132 size 48x16; Text 'BorderWidth'
   Bar "CornerRadius" at 560,10 size 40x120
   TextField "Label_CornerRadius" at 560,132 size 48x16; Text 'CornerRadius'
   Bar "CountSubDivisions" at 610,10 size 40x120
   TextField "Label_CountSubDivisions" at 610,132 size 48x16; Text 'CountSubDivisions'
   Bar "EdgeStyle" at 660,10 size 40x120
   TextField "Label_EdgeStyle" at 660,132 size 48x16; Text 'EdgeStyle'
   Bar "EdgeStyle_2" at 710,10 size 40x120
   TextField "Label_EdgeStyle_2" at 710,132 size 48x16; Text 'EdgeStyle_2'
   Bar "EdgeStyle_3" at 10,156 size 40x120
   TextField "Label_EdgeStyle_3" at 10,278 size 48x16; Text 'EdgeStyle_3'
   Bar "EdgeStyle_4" at 60,156 size 40x120
   TextField "Label_EdgeStyle_4" at 60,278 size 48x16; Text 'EdgeStyle_4'
   Bar "Flashing" at 110,156 size 40x120
   TextField "Label_Flashing" at 110,278 size 48x16; Text 'Flashing'
   Bar "FlashingOnLimitViolation" at 160,156 size 40x120
   TextField "Label_FlashingOnLimitViolation" at 160,278 size 48x16; Text 'FlashingOnLimitViolation'
   Bar "ForeColor" at 210,156 size 40x120
   TextField "Label_ForeColor" at 210,278 size 48x16; Text 'ForeColor'
   Bar "IntegerDigits" at 260,156 size 40x120
   TextField "Label_IntegerDigits" at 260,278 size 48x16; Text 'IntegerDigits'
   Bar "LargeTickLabelingStep" at 310,156 size 40x120
   TextField "Label_LargeTickLabelingStep" at 310,278 size 48x16; Text 'LargeTickLabelingStep'
   Bar "MaximumValue" at 360,156 size 40x120; MaximumValue 200
   TextField "Label_MaximumValue" at 360,278 size 48x16; Text 'MaximumValue'
   Bar "MinimumValue" at 410,156 size 40x120; MinimumValue -100
   TextField "Label_MinimumValue" at 410,278 size 48x16; Text 'MinimumValue'
   Bar "Precision" at 460,156 size 40x120
   TextField "Label_Precision" at 460,278 size 48x16; Text 'Precision'
   Bar "RangeLower1Color" at 510,156 size 40x120
   TextField "Label_RangeLower1Color" at 510,278 size 48x16; Text 'RangeLower1Color'
   Bar "RangeLower1Enabled" at 560,156 size 40x120
   TextField "Label_RangeLower1Enabled" at 560,278 size 48x16; Text 'RangeLower1Enabled'
   Bar "RangeLower2Color" at 610,156 size 40x120
   TextField "Label_RangeLower2Color" at 610,278 size 48x16; Text 'RangeLower2Color'
   Bar "RangeLower2Enabled" at 660,156 size 40x120
   TextField "Label_RangeLower2Enabled" at 660,278 size 48x16; Text 'RangeLower2Enabled'
   Bar "RangeNormalColor" at 710,156 size 40x120
   TextField "Label_RangeNormalColor" at 710,278 size 48x16; Text 'RangeNormalColor'
   Bar "RangeNormalEnabled" at 10,302 size 40x120
   TextField "Label_RangeNormalEnabled" at 10,424 size 48x16; Text 'RangeNormalEnabled'
   Bar "RangeUpper1Color" at 60,302 size 40x120
   TextField "Label_RangeUpper1Color" at 60,424 size 48x16; Text 'RangeUpper1Color'
   Bar "RangeUpper1Enabled" at 110,302 size 40x120
   TextField "Label_RangeUpper1Enabled" at 110,424 size 48x16; Text 'RangeUpper1Enabled'
   Bar "RangeUpper2Color" at 160,302 size 40x120
   TextField "Label_RangeUpper2Color" at 160,424 size 48x16; Text 'RangeUpper2Color'
   Bar "RangeUpper2Enabled" at 210,302 size 40x120
   TextField "Label_RangeUpper2Enabled" at 210,424 size 48x16; Text 'RangeUpper2Enabled'
   Bar "ScaleColor" at 260,302 size 40x120
   TextField "Label_ScaleColor" at 260,424 size 48x16; Text 'ScaleColor'
   Bar "ScaleGradation" at 310,302 size 40x120
   TextField "Label_ScaleGradation" at 310,424 size 48x16; Text 'ScaleGradation'
   Bar "ScaleLabelingDoubleLined" at 360,302 size 40x120
   TextField "Label_ScaleLabelingDoubleLined" at 360,424 size 48x16; Text 'ScaleLabelingDoubleLined'
   Bar "ScalePosition" at 410,302 size 40x120
   TextField "Label_ScalePosition" at 410,424 size 48x16; Text 'ScalePosition'
   Bar "SegmentColoring" at 460,302 size 40x120
   TextField "Label_SegmentColoring" at 460,424 size 48x16; Text 'SegmentColoring'
   Bar "ShowLimitLines" at 510,302 size 40x120
   TextField "Label_ShowLimitLines" at 510,424 size 48x16; Text 'ShowLimitLines'
   Bar "ShowLimitMarkers" at 560,302 size 40x120
   TextField "Label_ShowLimitMarkers" at 560,424 size 48x16; Text 'ShowLimitMarkers'
   Bar "ShowLimitRanges" at 610,302 size 40x120
   TextField "Label_ShowLimitRanges" at 610,424 size 48x16; Text 'ShowLimitRanges'
   Bar "ShowProcessValue" at 660,302 size 40x120
   TextField "Label_ShowProcessValue" at 660,424 size 48x16; Text 'ShowProcessValue'
   Bar "ShowScale" at 710,302 size 40x120
   TextField "Label_ShowScale" at 710,424 size 48x16; Text 'ShowScale'
   Button "Next" at 758,456 size 40x22; TextOff 'Text'
      on Click: ActivateScreen("P_Bar_2", 0)

screen "P_Bar_2" 800x480
   Bar "ShowTickLabels" at 10,10 size 40x120
   TextField "Label_ShowTickLabels" at 10,132 size 48x16; Text 'ShowTickLabels'
   Bar "Unit" at 60,10 size 40x120; Unit mm
   TextField "Label_Unit" at 60,132 size 48x16; Text 'Unit'
   Bar "UseAutoScaling" at 110,10 size 40x120
   TextField "Label_UseAutoScaling" at 110,132 size 48x16; Text 'UseAutoScaling'
   Bar "UseDesignColorSchema" at 160,10 size 40x120
   TextField "Label_UseDesignColorSchema" at 160,132 size 48x16; Text 'UseDesignColorSchema'
   Bar "UseExponentialFormat" at 210,10 size 40x120
   TextField "Label_UseExponentialFormat" at 210,132 size 48x16; Text 'UseExponentialFormat'
   Button "Next" at 758,456 size 40x22; TextOff 'Text'
      on Click: ActivateScreen("P_Switch_1", 0)

screen "P_Switch_1" 800x480
   Switch "Default" at 10,10 size 120x40; CaptionText 'Switch'; TextOff '0'; TextOn '1'
   TextField "Label_Default" at 10,52 size 128x16; Text 'Default'
   Switch "AboveUpperLimitColor" at 140,10 size 120x40; CaptionText 'Switch'; TextOff '0'; TextOn '1'
   TextField "Label_AboveUpperLimitColor" at 140,52 size 128x16; Text 'AboveUpperLimitColor'
   Switch "BackColor" at 270,10 size 120x40; CaptionText 'Switch'; TextOff '0'; TextOn '1'
   TextField "Label_BackColor" at 270,52 size 128x16; Text 'BackColor'
   Switch "BackFillStyle" at 400,10 size 120x40; CaptionText 'Switch'; TextOff '0'; TextOn '1'
   TextField "Label_BackFillStyle" at 400,52 size 128x16; Text 'BackFillStyle'
   Switch "BelowLowerLimitColor" at 530,10 size 120x40; CaptionText 'Switch'; TextOff '0'; TextOn '1'
   TextField "Label_BelowLowerLimitColor" at 530,52 size 128x16; Text 'BelowLowerLimitColor'
   Switch "BorderBackColor" at 660,10 size 120x40; CaptionText 'Switch'; TextOff '0'; TextOn '1'
   TextField "Label_BorderBackColor" at 660,52 size 128x16; Text 'BorderBackColor'
   Switch "BorderColor" at 10,76 size 120x40; CaptionText 'Switch'; TextOff '0'; TextOn '1'
   TextField "Label_BorderColor" at 10,118 size 128x16; Text 'BorderColor'
   Switch "BorderWidth" at 140,76 size 120x40; CaptionText 'Switch'; TextOff '0'; TextOn '1'
   TextField "Label_BorderWidth" at 140,118 size 128x16; Text 'BorderWidth'
   Switch "CaptionColor" at 270,76 size 120x40; CaptionText 'Switch'; TextOff '0'; TextOn '1'
   TextField "Label_CaptionColor" at 270,118 size 128x16; Text 'CaptionColor'
   Switch "CornerRadius" at 400,76 size 120x40; CaptionText 'Switch'; TextOff '0'; TextOn '1'
   TextField "Label_CornerRadius" at 400,118 size 128x16; Text 'CornerRadius'
   Switch "EdgeStyle" at 530,76 size 120x40; CaptionText 'Switch'; TextOff '0'; TextOn '1'
   TextField "Label_EdgeStyle" at 530,118 size 128x16; Text 'EdgeStyle'
   Switch "EdgeStyle_2" at 660,76 size 120x40; CaptionText 'Switch'; TextOff '0'; TextOn '1'
   TextField "Label_EdgeStyle_2" at 660,118 size 128x16; Text 'EdgeStyle_2'
   Switch "EdgeStyle_3" at 10,142 size 120x40; CaptionText 'Switch'; TextOff '0'; TextOn '1'
   TextField "Label_EdgeStyle_3" at 10,184 size 128x16; Text 'EdgeStyle_3'
   Switch "EdgeStyle_4" at 140,142 size 120x40; CaptionText 'Switch'; TextOff '0'; TextOn '1'
   TextField "Label_EdgeStyle_4" at 140,184 size 128x16; Text 'EdgeStyle_4'
   Switch "FirstGradientColor" at 270,142 size 120x40; CaptionText 'Switch'; TextOff '0'; TextOn '1'
   TextField "Label_FirstGradientColor" at 270,184 size 128x16; Text 'FirstGradientColor'
   Switch "FirstGradientOffset" at 400,142 size 120x40; CaptionText 'Switch'; TextOff '0'; TextOn '1'
   TextField "Label_FirstGradientOffset" at 400,184 size 128x16; Text 'FirstGradientOffset'
   Switch "FitToLargest" at 530,142 size 120x40; CaptionText 'Switch'; TextOff '0'; TextOn '1'
   TextField "Label_FitToLargest" at 530,184 size 128x16; Text 'FitToLargest'
   Switch "Flashing" at 660,142 size 120x40; CaptionText 'Switch'; TextOff '0'; TextOn '1'
   TextField "Label_Flashing" at 660,184 size 128x16; Text 'Flashing'
   Switch "FlashingOnLimitViolation" at 10,208 size 120x40; CaptionText 'Switch'; TextOff '0'; TextOn '1'
   TextField "Label_FlashingOnLimitViolation" at 10,250 size 128x16; Text 'FlashingOnLimitViolation'
   Switch "FocusColor" at 140,208 size 120x40; CaptionText 'Switch'; TextOff '0'; TextOn '1'
   TextField "Label_FocusColor" at 140,250 size 128x16; Text 'FocusColor'
   Switch "FocusWidth" at 270,208 size 120x40; CaptionText 'Switch'; TextOff '0'; TextOn '1'
   TextField "Label_FocusWidth" at 270,250 size 128x16; Text 'FocusWidth'
   Switch "ForeColor" at 400,208 size 120x40; CaptionText 'Switch'; TextOff '0'; TextOn '1'
   TextField "Label_ForeColor" at 400,250 size 128x16; Text 'ForeColor'
   Switch "HorizontalAlignment" at 530,208 size 120x40; CaptionText 'Switch'; TextOff '0'; TextOn '1'
   TextField "Label_HorizontalAlignment" at 530,250 size 128x16; Text 'HorizontalAlignment'
   Switch "HorizontalAlignment_2" at 660,208 size 120x40; CaptionText 'Switch'; TextOff '0'; TextOn '1'
   TextField "Label_HorizontalAlignment_2" at 660,250 size 128x16; Text 'HorizontalAlignment_2'
   Switch "HorizontalPictureAlignment" at 10,274 size 120x40; CaptionText 'Switch'; TextOff '0'; TextOn '1'
   TextField "Label_HorizontalPictureAlignment" at 10,316 size 128x16; Text 'HorizontalPictureAlignment'
   Switch "HorizontalPictureAlignment_2" at 140,274 size 120x40; CaptionText 'Switch'; TextOff '0'; TextOn '1'
   TextField "Label_HorizontalPictureAlignment_2" at 140,316 size 128x16; Text 'HorizontalPictureAlignment_2'
   Switch "InnerBackColorOff" at 270,274 size 120x40; CaptionText 'Switch'; TextOff '0'; TextOn '1'
   TextField "Label_InnerBackColorOff" at 270,316 size 128x16; Text 'InnerBackColorOff'
   Switch "InnerBackColorOn" at 400,274 size 120x40; CaptionText 'Switch'; TextOff '0'; TextOn '1'
   TextField "Label_InnerBackColorOn" at 400,316 size 128x16; Text 'InnerBackColorOn'
   Switch "MiddleGradientColor" at 530,274 size 120x40; CaptionText 'Switch'; TextOff '0'; TextOn '1'
   TextField "Label_MiddleGradientColor" at 530,316 size 128x16; Text 'MiddleGradientColor'
   Switch "PictureAreaBottomMargin" at 660,274 size 120x40; CaptionText 'Switch'; TextOff '0'; TextOn '1'
   TextField "Label_PictureAreaBottomMargin" at 660,316 size 128x16; Text 'PictureAreaBottomMargin'
   Switch "PictureAreaLeftMargin" at 10,340 size 120x40; CaptionText 'Switch'; TextOff '0'; TextOn '1'
   TextField "Label_PictureAreaLeftMargin" at 10,382 size 128x16; Text 'PictureAreaLeftMargin'
   Switch "PictureAreaRightMargin" at 140,340 size 120x40; CaptionText 'Switch'; TextOff '0'; TextOn '1'
   TextField "Label_PictureAreaRightMargin" at 140,382 size 128x16; Text 'PictureAreaRightMargin'
   Switch "PictureAreaTopMargin" at 270,340 size 120x40; CaptionText 'Switch'; TextOff '0'; TextOn '1'
   TextField "Label_PictureAreaTopMargin" at 270,382 size 128x16; Text 'PictureAreaTopMargin'
   Switch "SecondGradientColor" at 400,340 size 120x40; CaptionText 'Switch'; TextOff '0'; TextOn '1'
   TextField "Label_SecondGradientColor" at 400,382 size 128x16; Text 'SecondGradientColor'
   Switch "SecondGradientOffset" at 530,340 size 120x40; CaptionText 'Switch'; TextOff '0'; TextOn '1'
   TextField "Label_SecondGradientOffset" at 530,382 size 128x16; Text 'SecondGradientOffset'
   Switch "ShowCaption" at 660,340 size 120x40; CaptionText 'Switch'; TextOff '0'; TextOn '1'
   TextField "Label_ShowCaption" at 660,382 size 128x16; Text 'ShowCaption'
   Button "Next" at 758,456 size 40x22; TextOff 'Text'
      on Click: ActivateScreen("P_Switch_2", 0)

screen "P_Switch_2" 800x480
   Switch "SwitchOrientation" at 10,10 size 120x40; CaptionText 'Switch'; TextOff '0'; TextOn '1'
   TextField "Label_SwitchOrientation" at 10,52 size 128x16; Text 'SwitchOrientation'
   Switch "SwitchOrientation_2" at 140,10 size 120x40; CaptionText 'Switch'; TextOff '0'; TextOn '1'
   TextField "Label_SwitchOrientation_2" at 140,52 size 128x16; Text 'SwitchOrientation_2'
   Switch "SwitchOrientation_3" at 270,10 size 120x40; CaptionText 'Switch'; TextOff '0'; TextOn '1'
   TextField "Label_SwitchOrientation_3" at 270,52 size 128x16; Text 'SwitchOrientation_3'
   Switch "TextAreaBottomMargin" at 400,10 size 120x40; CaptionText 'Switch'; TextOff '0'; TextOn '1'
   TextField "Label_TextAreaBottomMargin" at 400,52 size 128x16; Text 'TextAreaBottomMargin'
   Switch "TextAreaLeftMargin" at 530,10 size 120x40; CaptionText 'Switch'; TextOff '0'; TextOn '1'
   TextField "Label_TextAreaLeftMargin" at 530,52 size 128x16; Text 'TextAreaLeftMargin'
   Switch "TextAreaRightMargin" at 660,10 size 120x40; CaptionText 'Switch'; TextOff '0'; TextOn '1'
   TextField "Label_TextAreaRightMargin" at 660,52 size 128x16; Text 'TextAreaRightMargin'
   Switch "TextAreaTopMargin" at 10,76 size 120x40; CaptionText 'Switch'; TextOff '0'; TextOn '1'
   TextField "Label_TextAreaTopMargin" at 10,118 size 128x16; Text 'TextAreaTopMargin'
   Switch "UseDesignColorSchema" at 140,76 size 120x40; CaptionText 'Switch'; TextOff '0'; TextOn '1'
   TextField "Label_UseDesignColorSchema" at 140,118 size 128x16; Text 'UseDesignColorSchema'
   Switch "UseFirstGradient" at 270,76 size 120x40; CaptionText 'Switch'; TextOff '0'; TextOn '1'
   TextField "Label_UseFirstGradient" at 270,118 size 128x16; Text 'UseFirstGradient'
   Switch "UseSecondGradient" at 400,76 size 120x40; CaptionText 'Switch'; TextOff '0'; TextOn '1'
   TextField "Label_UseSecondGradient" at 400,118 size 128x16; Text 'UseSecondGradient'
   Switch "VerticalAlignment" at 530,76 size 120x40; CaptionText 'Switch'; TextOff '0'; TextOn '1'
   TextField "Label_VerticalAlignment" at 530,118 size 128x16; Text 'VerticalAlignment'
   Switch "VerticalAlignment_2" at 660,76 size 120x40; CaptionText 'Switch'; TextOff '0'; TextOn '1'
   TextField "Label_VerticalAlignment_2" at 660,118 size 128x16; Text 'VerticalAlignment_2'
   Switch "VerticalPictureAlignment" at 10,142 size 120x40; CaptionText 'Switch'; TextOff '0'; TextOn '1'
   TextField "Label_VerticalPictureAlignment" at 10,184 size 128x16; Text 'VerticalPictureAlignment'
   Switch "VerticalPictureAlignment_2" at 140,142 size 120x40; CaptionText 'Switch'; TextOff '0'; TextOn '1'
   TextField "Label_VerticalPictureAlignment_2" at 140,184 size 128x16; Text 'VerticalPictureAlignment_2'
   Button "Next" at 758,456 size 40x22; TextOff 'Text'
      on Click: ActivateScreen("P_SymbolLibrary_1", 0)

screen "P_SymbolLibrary_1" 800x480
   SymbolLibrary "Default" at 10,10 size 60x60
   TextField "Label_Default" at 10,72 size 68x16; Text 'Default'
   SymbolLibrary "AboveUpperLimitColor" at 80,10 size 60x60
   TextField "Label_AboveUpperLimitColor" at 80,72 size 68x16; Text 'AboveUpperLimitColor'
   SymbolLibrary "BackColor" at 150,10 size 60x60
   TextField "Label_BackColor" at 150,72 size 68x16; Text 'BackColor'
   SymbolLibrary "BackFillStyle" at 220,10 size 60x60
   TextField "Label_BackFillStyle" at 220,72 size 68x16; Text 'BackFillStyle'
   SymbolLibrary "BelowLowerLimitColor" at 290,10 size 60x60
   TextField "Label_BelowLowerLimitColor" at 290,72 size 68x16; Text 'BelowLowerLimitColor'
   SymbolLibrary "BlinkColor" at 360,10 size 60x60
   TextField "Label_BlinkColor" at 360,72 size 68x16; Text 'BlinkColor'
   SymbolLibrary "FillColorMode" at 430,10 size 60x60
   TextField "Label_FillColorMode" at 430,72 size 68x16; Text 'FillColorMode'
   SymbolLibrary "FillColorMode_2" at 500,10 size 60x60
   TextField "Label_FillColorMode_2" at 500,72 size 68x16; Text 'FillColorMode_2'
   SymbolLibrary "FixedAspectRatio" at 570,10 size 60x60
   TextField "Label_FixedAspectRatio" at 570,72 size 68x16; Text 'FixedAspectRatio'
   SymbolLibrary "Flashing" at 640,10 size 60x60
   TextField "Label_Flashing" at 640,72 size 68x16; Text 'Flashing'
   SymbolLibrary "FlashingOnLimitViolation" at 710,10 size 60x60
   TextField "Label_FlashingOnLimitViolation" at 710,72 size 68x16; Text 'FlashingOnLimitViolation'
   SymbolLibrary "Flip" at 10,96 size 60x60
   TextField "Label_Flip" at 10,158 size 68x16; Text 'Flip'
   SymbolLibrary "Flip_2" at 80,96 size 60x60
   TextField "Label_Flip_2" at 80,158 size 68x16; Text 'Flip_2'
   SymbolLibrary "Flip_3" at 150,96 size 60x60
   TextField "Label_Flip_3" at 150,158 size 68x16; Text 'Flip_3'
   SymbolLibrary "ForeColor" at 220,96 size 60x60
   TextField "Label_ForeColor" at 220,158 size 68x16; Text 'ForeColor'
   SymbolLibrary "Rotation" at 290,96 size 60x60
   TextField "Label_Rotation" at 290,158 size 68x16; Text 'Rotation'
   SymbolLibrary "Rotation_2" at 360,96 size 60x60
   TextField "Label_Rotation_2" at 360,158 size 68x16; Text 'Rotation_2'
   SymbolLibrary "Rotation_3" at 430,96 size 60x60
   TextField "Label_Rotation_3" at 430,158 size 68x16; Text 'Rotation_3'
   Button "Next" at 758,456 size 40x22; TextOff 'Text'
      on Click: ActivateScreen("P_Slider_1", 0)

screen "P_Slider_1" 800x480
   Slider "Default" at 10,10 size 60x160; Caption 'SIMATIC'
   TextField "Label_Default" at 10,172 size 68x16; Text 'Default'
   Slider "BackColor" at 80,10 size 60x160; Caption 'SIMATIC'
   TextField "Label_BackColor" at 80,172 size 68x16; Text 'BackColor'
   Slider "BackFillStyle" at 150,10 size 60x160; Caption 'SIMATIC'
   TextField "Label_BackFillStyle" at 150,172 size 68x16; Text 'BackFillStyle'
   Slider "BarBackColor" at 220,10 size 60x160; Caption 'SIMATIC'
   TextField "Label_BarBackColor" at 220,172 size 68x16; Text 'BarBackColor'
   Slider "BarColor" at 290,10 size 60x160; Caption 'SIMATIC'
   TextField "Label_BarColor" at 290,172 size 68x16; Text 'BarColor'
   Slider "BarOrientation" at 360,10 size 60x160; Caption 'SIMATIC'
   TextField "Label_BarOrientation" at 360,172 size 68x16; Text 'BarOrientation'
   Slider "BarOrientation_2" at 430,10 size 60x160; Caption 'SIMATIC'
   TextField "Label_BarOrientation_2" at 430,172 size 68x16; Text 'BarOrientation_2'
   Slider "BarOrientation_3" at 500,10 size 60x160; Caption 'SIMATIC'
   TextField "Label_BarOrientation_3" at 500,172 size 68x16; Text 'BarOrientation_3'
   Slider "BorderBackColor" at 570,10 size 60x160; Caption 'SIMATIC'
   TextField "Label_BorderBackColor" at 570,172 size 68x16; Text 'BorderBackColor'
   Slider "BorderBrightColor3D" at 640,10 size 60x160; Caption 'SIMATIC'
   TextField "Label_BorderBrightColor3D" at 640,172 size 68x16; Text 'BorderBrightColor3D'
   Slider "BorderColor" at 710,10 size 60x160; Caption 'SIMATIC'
   TextField "Label_BorderColor" at 710,172 size 68x16; Text 'BorderColor'
   Slider "BorderInnerStyle3D" at 10,196 size 60x160; Caption 'SIMATIC'
   TextField "Label_BorderInnerStyle3D" at 10,358 size 68x16; Text 'BorderInnerStyle3D'
   Slider "BorderInnerStyle3D_2" at 80,196 size 60x160; Caption 'SIMATIC'
   TextField "Label_BorderInnerStyle3D_2" at 80,358 size 68x16; Text 'BorderInnerStyle3D_2'
   Slider "BorderInnerWidth3D" at 150,196 size 60x160; Caption 'SIMATIC'
   TextField "Label_BorderInnerWidth3D" at 150,358 size 68x16; Text 'BorderInnerWidth3D'
   Slider "BorderOuterStyle3D" at 220,196 size 60x160; Caption 'SIMATIC'
   TextField "Label_BorderOuterStyle3D" at 220,358 size 68x16; Text 'BorderOuterStyle3D'
   Slider "BorderOuterStyle3D_2" at 290,196 size 60x160; Caption 'SIMATIC'
   TextField "Label_BorderOuterStyle3D_2" at 290,358 size 68x16; Text 'BorderOuterStyle3D_2'
   Slider "BorderOuterWidth3D" at 360,196 size 60x160; Caption 'SIMATIC'
   TextField "Label_BorderOuterWidth3D" at 360,358 size 68x16; Text 'BorderOuterWidth3D'
   Slider "BorderShadeColor3D" at 430,196 size 60x160; Caption 'SIMATIC'
   TextField "Label_BorderShadeColor3D" at 430,358 size 68x16; Text 'BorderShadeColor3D'
   Slider "BorderWidth" at 500,196 size 60x160; Caption 'SIMATIC'
   TextField "Label_BorderWidth" at 500,358 size 68x16; Text 'BorderWidth'
   Slider "CornerRadius" at 570,196 size 60x160; Caption 'SIMATIC'
   TextField "Label_CornerRadius" at 570,358 size 68x16; Text 'CornerRadius'
   Slider "EdgeStyle" at 640,196 size 60x160; Caption 'SIMATIC'
   TextField "Label_EdgeStyle" at 640,358 size 68x16; Text 'EdgeStyle'
   Slider "EdgeStyle_2" at 710,196 size 60x160; Caption 'SIMATIC'
   TextField "Label_EdgeStyle_2" at 710,358 size 68x16; Text 'EdgeStyle_2'
   Button "Next" at 758,456 size 40x22; TextOff 'Text'
      on Click: ActivateScreen("P_Slider_2", 0)

screen "P_Slider_2" 800x480
   Slider "EdgeStyle_3" at 10,10 size 60x160; Caption 'SIMATIC'
   TextField "Label_EdgeStyle_3" at 10,172 size 68x16; Text 'EdgeStyle_3'
   Slider "EdgeStyle_4" at 80,10 size 60x160; Caption 'SIMATIC'
   TextField "Label_EdgeStyle_4" at 80,172 size 68x16; Text 'EdgeStyle_4'
   Slider "Flashing" at 150,10 size 60x160; Caption 'SIMATIC'
   TextField "Label_Flashing" at 150,172 size 68x16; Text 'Flashing'
   Slider "FocusColor" at 220,10 size 60x160; Caption 'SIMATIC'
   TextField "Label_FocusColor" at 220,172 size 68x16; Text 'FocusColor'
   Slider "FocusWidth" at 290,10 size 60x160; Caption 'SIMATIC'
   TextField "Label_FocusWidth" at 290,172 size 68x16; Text 'FocusWidth'
   Slider "ForeColor" at 360,10 size 60x160; Caption 'SIMATIC'
   TextField "Label_ForeColor" at 360,172 size 68x16; Text 'ForeColor'
   Slider "LabelColor" at 430,10 size 60x160; Caption 'SIMATIC'
   TextField "Label_LabelColor" at 430,172 size 68x16; Text 'LabelColor'
   Slider "MaximumValue" at 500,10 size 60x160; Caption 'SIMATIC'
   TextField "Label_MaximumValue" at 500,172 size 68x16; Text 'MaximumValue'
   Slider "MinimumValue" at 570,10 size 60x160; Caption 'SIMATIC'
   TextField "Label_MinimumValue" at 570,172 size 68x16; Text 'MinimumValue'
   Slider "RangeLower1Color" at 640,10 size 60x160; Caption 'SIMATIC'
   TextField "Label_RangeLower1Color" at 640,172 size 68x16; Text 'RangeLower1Color'
   Slider "RangeLower1Enabled" at 710,10 size 60x160; Caption 'SIMATIC'
   TextField "Label_RangeLower1Enabled" at 710,172 size 68x16; Text 'RangeLower1Enabled'
   Slider "RangeLower2Color" at 10,196 size 60x160; Caption 'SIMATIC'
   TextField "Label_RangeLower2Color" at 10,358 size 68x16; Text 'RangeLower2Color'
   Slider "RangeLower2Enabled" at 80,196 size 60x160; Caption 'SIMATIC'
   TextField "Label_RangeLower2Enabled" at 80,358 size 68x16; Text 'RangeLower2Enabled'
   Slider "RangeNormalColor" at 150,196 size 60x160; Caption 'SIMATIC'
   TextField "Label_RangeNormalColor" at 150,358 size 68x16; Text 'RangeNormalColor'
   Slider "RangeNormalEnabled" at 220,196 size 60x160; Caption 'SIMATIC'
   TextField "Label_RangeNormalEnabled" at 220,358 size 68x16; Text 'RangeNormalEnabled'
   Slider "RangeUpper1Color" at 290,196 size 60x160; Caption 'SIMATIC'
   TextField "Label_RangeUpper1Color" at 290,358 size 68x16; Text 'RangeUpper1Color'
   Slider "RangeUpper1Enabled" at 360,196 size 60x160; Caption 'SIMATIC'
   TextField "Label_RangeUpper1Enabled" at 360,358 size 68x16; Text 'RangeUpper1Enabled'
   Slider "RangeUpper2Color" at 430,196 size 60x160; Caption 'SIMATIC'
   TextField "Label_RangeUpper2Color" at 430,358 size 68x16; Text 'RangeUpper2Color'
   Slider "RangeUpper2Enabled" at 500,196 size 60x160; Caption 'SIMATIC'
   TextField "Label_RangeUpper2Enabled" at 500,358 size 68x16; Text 'RangeUpper2Enabled'
   Slider "ScalePosition" at 570,196 size 60x160; Caption 'SIMATIC'
   TextField "Label_ScalePosition" at 570,358 size 68x16; Text 'ScalePosition'
   Slider "ShowBar" at 640,196 size 60x160; Caption 'SIMATIC'
   TextField "Label_ShowBar" at 640,358 size 68x16; Text 'ShowBar'
   Slider "ShowLimitLines" at 710,196 size 60x160; Caption 'SIMATIC'
   TextField "Label_ShowLimitLines" at 710,358 size 68x16; Text 'ShowLimitLines'
   Button "Next" at 758,456 size 40x22; TextOff 'Text'
      on Click: ActivateScreen("P_Slider_3", 0)

screen "P_Slider_3" 800x480
   Slider "ShowLimitMarkers" at 10,10 size 60x160; Caption 'SIMATIC'
   TextField "Label_ShowLimitMarkers" at 10,172 size 68x16; Text 'ShowLimitMarkers'
   Slider "ShowLimitRanges" at 80,10 size 60x160; Caption 'SIMATIC'
   TextField "Label_ShowLimitRanges" at 80,172 size 68x16; Text 'ShowLimitRanges'
   Slider "ShowPosition" at 150,10 size 60x160; Caption 'SIMATIC'
   TextField "Label_ShowPosition" at 150,172 size 68x16; Text 'ShowPosition'
   Slider "ShowScale" at 220,10 size 60x160; Caption 'SIMATIC'
   TextField "Label_ShowScale" at 220,172 size 68x16; Text 'ShowScale'
   Slider "ShowThumb" at 290,10 size 60x160; Caption 'SIMATIC'
   TextField "Label_ShowThumb" at 290,172 size 68x16; Text 'ShowThumb'
   Slider "ShowTickLabels" at 360,10 size 60x160; Caption 'SIMATIC'
   TextField "Label_ShowTickLabels" at 360,172 size 68x16; Text 'ShowTickLabels'
   Slider "ShowTicks" at 430,10 size 60x160; Caption 'SIMATIC'
   TextField "Label_ShowTicks" at 430,172 size 68x16; Text 'ShowTicks'
   Slider "ThumbBackColor" at 500,10 size 60x160; Caption 'SIMATIC'
   TextField "Label_ThumbBackColor" at 500,172 size 68x16; Text 'ThumbBackColor'
   Slider "UseDesignColorSchema" at 570,10 size 60x160; Caption 'SIMATIC'
   TextField "Label_UseDesignColorSchema" at 570,172 size 68x16; Text 'UseDesignColorSchema'
   Button "Next" at 758,456 size 40x22; TextOff 'Text'
      on Click: ActivateScreen("P_Gauge_1", 0)

screen "P_Gauge_1" 800x480
   Gauge "Default" at 10,10 size 150x150; CaptionText 'SIMATIC'
   TextField "Label_Default" at 10,162 size 158x16; Text 'Default'
   Gauge "AngleMax" at 170,10 size 150x150; CaptionText 'SIMATIC'
   TextField "Label_AngleMax" at 170,162 size 158x16; Text 'AngleMax'
   Gauge "AngleMin" at 330,10 size 150x150; CaptionText 'SIMATIC'
   TextField "Label_AngleMin" at 330,162 size 158x16; Text 'AngleMin'
   Gauge "BackColor" at 490,10 size 150x150; CaptionText 'SIMATIC'
   TextField "Label_BackColor" at 490,162 size 158x16; Text 'BackColor'
   Gauge "BackFillStyle" at 10,186 size 150x150; CaptionText 'SIMATIC'
   TextField "Label_BackFillStyle" at 10,338 size 158x16; Text 'BackFillStyle'
   Gauge "BorderBackColor" at 170,186 size 150x150; CaptionText 'SIMATIC'
   TextField "Label_BorderBackColor" at 170,338 size 158x16; Text 'BorderBackColor'
   Gauge "BorderColor" at 330,186 size 150x150; CaptionText 'SIMATIC'
   TextField "Label_BorderColor" at 330,338 size 158x16; Text 'BorderColor'
   Gauge "BorderWidth" at 490,186 size 150x150; CaptionText 'SIMATIC'
   TextField "Label_BorderWidth" at 490,338 size 158x16; Text 'BorderWidth'
   Button "Next" at 758,456 size 40x22; TextOff 'Text'
      on Click: ActivateScreen("P_Gauge_2", 0)

screen "P_Gauge_2" 800x480
   Gauge "CaptionColor" at 10,10 size 150x150; CaptionText 'SIMATIC'
   TextField "Label_CaptionColor" at 10,162 size 158x16; Text 'CaptionColor'
   Gauge "CaptionTop" at 170,10 size 150x150; CaptionText 'SIMATIC'
   TextField "Label_CaptionTop" at 170,162 size 158x16; Text 'CaptionTop'
   Gauge "CenterColor" at 330,10 size 150x150; CaptionText 'SIMATIC'
   TextField "Label_CenterColor" at 330,162 size 158x16; Text 'CenterColor'
   Gauge "CenterSize" at 490,10 size 150x150; CaptionText 'SIMATIC'
   TextField "Label_CenterSize" at 490,162 size 158x16; Text 'CenterSize'
   Gauge "CornerRadius" at 10,186 size 150x150; CaptionText 'SIMATIC'
   TextField "Label_CornerRadius" at 10,338 size 158x16; Text 'CornerRadius'
   Gauge "DialColor" at 170,186 size 150x150; CaptionText 'SIMATIC'
   TextField "Label_DialColor" at 170,338 size 158x16; Text 'DialColor'
   Gauge "DialFillStyle" at 330,186 size 150x150; CaptionText 'SIMATIC'
   TextField "Label_DialFillStyle" at 330,338 size 158x16; Text 'DialFillStyle'
   Gauge "DialSize" at 490,186 size 150x150; CaptionText 'SIMATIC'
   TextField "Label_DialSize" at 490,338 size 158x16; Text 'DialSize'
   Button "Next" at 758,456 size 40x22; TextOff 'Text'
      on Click: ActivateScreen("P_Gauge_3", 0)

screen "P_Gauge_3" 800x480
   Gauge "EdgeStyle" at 10,10 size 150x150; CaptionText 'SIMATIC'
   TextField "Label_EdgeStyle" at 10,162 size 158x16; Text 'EdgeStyle'
   Gauge "EdgeStyle_2" at 170,10 size 150x150; CaptionText 'SIMATIC'
   TextField "Label_EdgeStyle_2" at 170,162 size 158x16; Text 'EdgeStyle_2'
   Gauge "EdgeStyle_3" at 330,10 size 150x150; CaptionText 'SIMATIC'
   TextField "Label_EdgeStyle_3" at 330,162 size 158x16; Text 'EdgeStyle_3'
   Gauge "EdgeStyle_4" at 490,10 size 150x150; CaptionText 'SIMATIC'
   TextField "Label_EdgeStyle_4" at 490,162 size 158x16; Text 'EdgeStyle_4'
   Gauge "Gradation" at 10,186 size 150x150; CaptionText 'SIMATIC'
   TextField "Label_Gradation" at 10,338 size 158x16; Text 'Gradation'
   Gauge "InnerDialColor" at 170,186 size 150x150; CaptionText 'SIMATIC'
   TextField "Label_InnerDialColor" at 170,338 size 158x16; Text 'InnerDialColor'
   Gauge "InnerDialInnerDistance" at 330,186 size 150x150; CaptionText 'SIMATIC'
   TextField "Label_InnerDialInnerDistance" at 330,338 size 158x16; Text 'InnerDialInnerDistance'
   Gauge "InnerDialOuterDistance" at 490,186 size 150x150; CaptionText 'SIMATIC'
   TextField "Label_InnerDialOuterDistance" at 490,338 size 158x16; Text 'InnerDialOuterDistance'
   Button "Next" at 758,456 size 40x22; TextOff 'Text'
      on Click: ActivateScreen("P_Gauge_4", 0)

screen "P_Gauge_4" 800x480
   Gauge "LockSquaredExtent" at 10,10 size 150x150; CaptionText 'SIMATIC'
   TextField "Label_LockSquaredExtent" at 10,162 size 158x16; Text 'LockSquaredExtent'
   Gauge "MaximumValue" at 170,10 size 150x150; CaptionText 'SIMATIC'
   TextField "Label_MaximumValue" at 170,162 size 158x16; Text 'MaximumValue'
   Gauge "MinimumValue" at 330,10 size 150x150; CaptionText 'SIMATIC'
   TextField "Label_MinimumValue" at 330,162 size 158x16; Text 'MinimumValue'
   Gauge "NeedleHeight" at 490,10 size 150x150; CaptionText 'SIMATIC'
   TextField "Label_NeedleHeight" at 490,162 size 158x16; Text 'NeedleHeight'
   Gauge "PointerColor" at 10,186 size 150x150; CaptionText 'SIMATIC'
   TextField "Label_PointerColor" at 10,338 size 158x16; Text 'PointerColor'
   Gauge "RangeLower1Color" at 170,186 size 150x150; CaptionText 'SIMATIC'
   TextField "Label_RangeLower1Color" at 170,338 size 158x16; Text 'RangeLower1Color'
   Gauge "RangeLower1Enabled" at 330,186 size 150x150; CaptionText 'SIMATIC'
   TextField "Label_RangeLower1Enabled" at 330,338 size 158x16; Text 'RangeLower1Enabled'
   Gauge "RangeLower2Color" at 490,186 size 150x150; CaptionText 'SIMATIC'
   TextField "Label_RangeLower2Color" at 490,338 size 158x16; Text 'RangeLower2Color'
   Button "Next" at 758,456 size 40x22; TextOff 'Text'
      on Click: ActivateScreen("P_Gauge_5", 0)

screen "P_Gauge_5" 800x480
   Gauge "RangeLower2Enabled" at 10,10 size 150x150; CaptionText 'SIMATIC'
   TextField "Label_RangeLower2Enabled" at 10,162 size 158x16; Text 'RangeLower2Enabled'
   Gauge "RangeNormalColor" at 170,10 size 150x150; CaptionText 'SIMATIC'
   TextField "Label_RangeNormalColor" at 170,162 size 158x16; Text 'RangeNormalColor'
   Gauge "RangeNormalEnabled" at 330,10 size 150x150; CaptionText 'SIMATIC'
   TextField "Label_RangeNormalEnabled" at 330,162 size 158x16; Text 'RangeNormalEnabled'
   Gauge "RangeUpper1Color" at 490,10 size 150x150; CaptionText 'SIMATIC'
   TextField "Label_RangeUpper1Color" at 490,162 size 158x16; Text 'RangeUpper1Color'
   Gauge "RangeUpper1Enabled" at 10,186 size 150x150; CaptionText 'SIMATIC'
   TextField "Label_RangeUpper1Enabled" at 10,338 size 158x16; Text 'RangeUpper1Enabled'
   Gauge "RangeUpper1Start" at 170,186 size 150x150; CaptionText 'SIMATIC'
   TextField "Label_RangeUpper1Start" at 170,338 size 158x16; Text 'RangeUpper1Start'
   Gauge "RangeUpper2Color" at 330,186 size 150x150; CaptionText 'SIMATIC'
   TextField "Label_RangeUpper2Color" at 330,338 size 158x16; Text 'RangeUpper2Color'
   Gauge "RangeUpper2Enabled" at 490,186 size 150x150; CaptionText 'SIMATIC'
   TextField "Label_RangeUpper2Enabled" at 490,338 size 158x16; Text 'RangeUpper2Enabled'
   Button "Next" at 758,456 size 40x22; TextOff 'Text'
      on Click: ActivateScreen("P_Gauge_6", 0)

screen "P_Gauge_6" 800x480
   Gauge "RangeUpper2Start" at 10,10 size 150x150; CaptionText 'SIMATIC'
   TextField "Label_RangeUpper2Start" at 10,162 size 158x16; Text 'RangeUpper2Start'
   Gauge "ScaleLabelColor" at 170,10 size 150x150; CaptionText 'SIMATIC'
   TextField "Label_ScaleLabelColor" at 170,162 size 158x16; Text 'ScaleLabelColor'
   Gauge "ScaleTickColor" at 330,10 size 150x150; CaptionText 'SIMATIC'
   TextField "Label_ScaleTickColor" at 330,162 size 158x16; Text 'ScaleTickColor'
   Gauge "ScaleTickLabelPosition" at 490,10 size 150x150; CaptionText 'SIMATIC'
   TextField "Label_ScaleTickLabelPosition" at 490,162 size 158x16; Text 'ScaleTickLabelPosition'
   Gauge "ScaleTickLength" at 10,186 size 150x150; CaptionText 'SIMATIC'
   TextField "Label_ScaleTickLength" at 10,338 size 158x16; Text 'ScaleTickLength'
   Gauge "ScaleTickPosition" at 170,186 size 150x150; CaptionText 'SIMATIC'
   TextField "Label_ScaleTickPosition" at 170,338 size 158x16; Text 'ScaleTickPosition'
   Gauge "ShowDecimalPoint" at 330,186 size 150x150; CaptionText 'SIMATIC'
   TextField "Label_ShowDecimalPoint" at 330,338 size 158x16; Text 'ShowDecimalPoint'
   Gauge "ShowInnerDial" at 490,186 size 150x150; CaptionText 'SIMATIC'
   TextField "Label_ShowInnerDial" at 490,338 size 158x16; Text 'ShowInnerDial'
   Button "Next" at 758,456 size 40x22; TextOff 'Text'
      on Click: ActivateScreen("P_Gauge_7", 0)

screen "P_Gauge_7" 800x480
   Gauge "ShowLimitRanges" at 10,10 size 150x150; CaptionText 'SIMATIC'
   TextField "Label_ShowLimitRanges" at 10,162 size 158x16; Text 'ShowLimitRanges'
   Gauge "ShowPeakValuePointer" at 170,10 size 150x150; CaptionText 'SIMATIC'
   TextField "Label_ShowPeakValuePointer" at 170,162 size 158x16; Text 'ShowPeakValuePointer'
   Gauge "UnitColor" at 330,10 size 150x150; CaptionText 'SIMATIC'
   TextField "Label_UnitColor" at 330,162 size 158x16; Text 'UnitColor'
   Gauge "UnitTop" at 490,10 size 150x150; CaptionText 'SIMATIC'
   TextField "Label_UnitTop" at 490,162 size 158x16; Text 'UnitTop'
   Gauge "UseDesignColorSchema" at 10,186 size 150x150; CaptionText 'SIMATIC'
   TextField "Label_UseDesignColorSchema" at 10,338 size 158x16; Text 'UseDesignColorSchema'
   Button "Next" at 758,456 size 40x22; TextOff 'Text'
      on Click: ActivateScreen("P_Clock_1", 0)

screen "P_Clock_1" 800x480
   Clock "Default" at 10,10 size 150x150
   TextField "Label_Default" at 10,162 size 158x16; Text 'Default'
   Clock "Analog" at 170,10 size 150x150
   TextField "Label_Analog" at 170,162 size 158x16; Text 'Analog'
   Clock "BackFillStyle" at 330,10 size 150x150
   TextField "Label_BackFillStyle" at 330,162 size 158x16; Text 'BackFillStyle'
   Clock "BorderBackColor" at 490,10 size 150x150
   TextField "Label_BorderBackColor" at 490,162 size 158x16; Text 'BorderBackColor'
   Clock "BorderColor" at 10,186 size 150x150
   TextField "Label_BorderColor" at 10,338 size 158x16; Text 'BorderColor'
   Clock "BorderWidth" at 170,186 size 150x150
   TextField "Label_BorderWidth" at 170,338 size 158x16; Text 'BorderWidth'
   Clock "CornerRadius" at 330,186 size 150x150
   TextField "Label_CornerRadius" at 330,338 size 158x16; Text 'CornerRadius'
   Clock "DialColor" at 490,186 size 150x150
   TextField "Label_DialColor" at 490,338 size 158x16; Text 'DialColor'
   Button "Next" at 758,456 size 40x22; TextOff 'Text'
      on Click: ActivateScreen("P_Clock_2", 0)

screen "P_Clock_2" 800x480
   Clock "EdgeStyle" at 10,10 size 150x150
   TextField "Label_EdgeStyle" at 10,162 size 158x16; Text 'EdgeStyle'
   Clock "EdgeStyle_2" at 170,10 size 150x150
   TextField "Label_EdgeStyle_2" at 170,162 size 158x16; Text 'EdgeStyle_2'
   Clock "EdgeStyle_3" at 330,10 size 150x150
   TextField "Label_EdgeStyle_3" at 330,162 size 158x16; Text 'EdgeStyle_3'
   Clock "EdgeStyle_4" at 490,10 size 150x150
   TextField "Label_EdgeStyle_4" at 490,162 size 158x16; Text 'EdgeStyle_4'
   Clock "Flashing" at 10,186 size 150x150
   TextField "Label_Flashing" at 10,338 size 158x16; Text 'Flashing'
   Clock "HourNeedleHeight" at 170,186 size 150x150
   TextField "Label_HourNeedleHeight" at 170,338 size 158x16; Text 'HourNeedleHeight'
   Clock "HourNeedleWidth" at 330,186 size 150x150
   TextField "Label_HourNeedleWidth" at 330,338 size 158x16; Text 'HourNeedleWidth'
   Clock "LockSquaredExtent" at 490,186 size 150x150
   TextField "Label_LockSquaredExtent" at 490,338 size 158x16; Text 'LockSquaredExtent'
   Button "Next" at 758,456 size 40x22; TextOff 'Text'
      on Click: ActivateScreen("P_Clock_3", 0)

screen "P_Clock_3" 800x480
   Clock "MinuteNeedleHeight" at 10,10 size 150x150
   TextField "Label_MinuteNeedleHeight" at 10,162 size 158x16; Text 'MinuteNeedleHeight'
   Clock "MinuteNeedleWidth" at 170,10 size 150x150
   TextField "Label_MinuteNeedleWidth" at 170,162 size 158x16; Text 'MinuteNeedleWidth'
   Clock "NeedleBorderColor" at 330,10 size 150x150
   TextField "Label_NeedleBorderColor" at 330,162 size 158x16; Text 'NeedleBorderColor'
   Clock "NeedleColor" at 490,10 size 150x150
   TextField "Label_NeedleColor" at 490,162 size 158x16; Text 'NeedleColor'
   Clock "NeedleFillStyle" at 10,186 size 150x150
   TextField "Label_NeedleFillStyle" at 10,338 size 158x16; Text 'NeedleFillStyle'
   Clock "NumberStyle" at 170,186 size 150x150
   TextField "Label_NumberStyle" at 170,338 size 158x16; Text 'NumberStyle'
   Clock "NumberStyle_2" at 330,186 size 150x150
   TextField "Label_NumberStyle_2" at 330,338 size 158x16; Text 'NumberStyle_2'
   Clock "SecondNeedleHeight" at 490,186 size 150x150
   TextField "Label_SecondNeedleHeight" at 490,338 size 158x16; Text 'SecondNeedleHeight'
   Button "Next" at 758,456 size 40x22; TextOff 'Text'
      on Click: ActivateScreen("P_Clock_4", 0)

screen "P_Clock_4" 800x480
   Clock "SecondNeedleWidth" at 10,10 size 150x150
   TextField "Label_SecondNeedleWidth" at 10,162 size 158x16; Text 'SecondNeedleWidth'
   Clock "ShowTicks" at 170,10 size 150x150
   TextField "Label_ShowTicks" at 170,162 size 158x16; Text 'ShowTicks'
   Clock "TickDistance" at 330,10 size 150x150
   TextField "Label_TickDistance" at 330,162 size 158x16; Text 'TickDistance'
   Clock "TickStyle" at 490,10 size 150x150
   TextField "Label_TickStyle" at 490,162 size 158x16; Text 'TickStyle'
   Clock "TicksColor" at 10,186 size 150x150
   TextField "Label_TicksColor" at 10,338 size 158x16; Text 'TicksColor'
   Clock "UseDesignColorSchema" at 170,186 size 150x150
   TextField "Label_UseDesignColorSchema" at 170,338 size 158x16; Text 'UseDesignColorSchema'
   Button "Next" at 758,456 size 40x22; TextOff 'Text'
      on Click: ActivateScreen("P_Line_1", 0)

screen "P_IOField_1" 800x480
   IOField "Default" at 10,10 size 100x30
   TextField "Label_Default" at 10,42 size 108x16; Text 'Default'
   IOField "AboveUpperLimitColor" at 120,10 size 100x30
   TextField "Label_AboveUpperLimitColor" at 120,42 size 108x16; Text 'AboveUpperLimitColor'
   IOField "BackColor" at 230,10 size 100x30
   TextField "Label_BackColor" at 230,42 size 108x16; Text 'BackColor'
   IOField "BackFillStyle" at 340,10 size 100x30
   TextField "Label_BackFillStyle" at 340,42 size 108x16; Text 'BackFillStyle'
   IOField "BelowLowerLimitColor" at 450,10 size 100x30
   TextField "Label_BelowLowerLimitColor" at 450,42 size 108x16; Text 'BelowLowerLimitColor'
   IOField "BorderBackColor" at 560,10 size 100x30
   TextField "Label_BorderBackColor" at 560,42 size 108x16; Text 'BorderBackColor'
   IOField "BorderColor" at 670,10 size 100x30
   TextField "Label_BorderColor" at 670,42 size 108x16; Text 'BorderColor'
   IOField "BorderWidth" at 10,66 size 100x30
   TextField "Label_BorderWidth" at 10,98 size 108x16; Text 'BorderWidth'
   IOField "BottomMargin" at 120,66 size 100x30
   TextField "Label_BottomMargin" at 120,98 size 108x16; Text 'BottomMargin'
   IOField "CornerRadius" at 230,66 size 100x30
   TextField "Label_CornerRadius" at 230,98 size 108x16; Text 'CornerRadius'
   IOField "DataFormat_3" at 340,66 size 100x30
   TextField "Label_DataFormat_3" at 340,98 size 108x16; Text 'DataFormat_3'
   IOField "EdgeStyle" at 450,66 size 100x30
   TextField "Label_EdgeStyle" at 450,98 size 108x16; Text 'EdgeStyle'
   IOField "EdgeStyle_2" at 560,66 size 100x30
   TextField "Label_EdgeStyle_2" at 560,98 size 108x16; Text 'EdgeStyle_2'
   IOField "EdgeStyle_3" at 670,66 size 100x30
   TextField "Label_EdgeStyle_3" at 670,98 size 108x16; Text 'EdgeStyle_3'
   IOField "EdgeStyle_4" at 10,122 size 100x30
   TextField "Label_EdgeStyle_4" at 10,154 size 108x16; Text 'EdgeStyle_4'
   IOField "FieldLength" at 120,122 size 100x30
   TextField "Label_FieldLength" at 120,154 size 108x16; Text 'FieldLength'
   IOField "FitToLargest" at 230,122 size 100x30
   TextField "Label_FitToLargest" at 230,154 size 108x16; Text 'FitToLargest'
   IOField "Flashing" at 340,122 size 100x30
   TextField "Label_Flashing" at 340,154 size 108x16; Text 'Flashing'
   IOField "ForeColor" at 450,122 size 100x30
   TextField "Label_ForeColor" at 450,154 size 108x16; Text 'ForeColor'
   IOField "FormatPattern" at 560,122 size 100x30; FormatPattern 99.9
   TextField "Label_FormatPattern" at 560,154 size 108x16; Text 'FormatPattern'
   IOField "HorizontalAlignment" at 670,122 size 100x30
   TextField "Label_HorizontalAlignment" at 670,154 size 108x16; Text 'HorizontalAlignment'
   IOField "HorizontalAlignment_2" at 10,178 size 100x30
   TextField "Label_HorizontalAlignment_2" at 10,210 size 108x16; Text 'HorizontalAlignment_2'
   IOField "LeftMargin" at 120,178 size 100x30
   TextField "Label_LeftMargin" at 120,210 size 108x16; Text 'LeftMargin'
   IOField "Mode" at 230,178 size 100x30
   TextField "Label_Mode" at 230,210 size 108x16; Text 'Mode'
   IOField "Mode_2" at 340,178 size 100x30
   TextField "Label_Mode_2" at 340,210 size 108x16; Text 'Mode_2'
   IOField "RightMargin" at 450,178 size 100x30
   TextField "Label_RightMargin" at 450,210 size 108x16; Text 'RightMargin'
   IOField "ShiftDecimalPoint" at 560,178 size 100x30
   TextField "Label_ShiftDecimalPoint" at 560,210 size 108x16; Text 'ShiftDecimalPoint'
   IOField "ShowLeadingZeros" at 670,178 size 100x30
   TextField "Label_ShowLeadingZeros" at 670,210 size 108x16; Text 'ShowLeadingZeros'
   IOField "TopMargin" at 10,234 size 100x30
   TextField "Label_TopMargin" at 10,266 size 108x16; Text 'TopMargin'
   IOField "Unit" at 120,234 size 100x30; Unit mm
   TextField "Label_Unit" at 120,266 size 108x16; Text 'Unit'
   IOField "UseDesignColorSchema" at 230,234 size 100x30
   TextField "Label_UseDesignColorSchema" at 230,266 size 108x16; Text 'UseDesignColorSchema'
   IOField "VerticalAlignment" at 340,234 size 100x30
   TextField "Label_VerticalAlignment" at 340,266 size 108x16; Text 'VerticalAlignment'
   IOField "VerticalAlignment_2" at 450,234 size 100x30
   TextField "Label_VerticalAlignment_2" at 450,266 size 108x16; Text 'VerticalAlignment_2'
   Button "Next" at 758,456 size 40x22; TextOff 'Text'
      on Click: ActivateScreen("P_Button_1", 0)

screen "D_Button_1" 800x480
   Button "Static" at 6,4 size 100x40; TextOff 'Text'
   TextField "Label_Static" at 6,76 size 148x16; Text 'Static'
   Button "A_Range" at 158,4 size 100x40; TextOff 'Text'
      Appearance <- "D_Range"
   TextField "Label_A_Range" at 158,76 size 148x16; Text 'A_Range'
   Button "A_Flash" at 310,4 size 100x40; TextOff 'Text'
      Appearance <- "D_Range"
   TextField "Label_A_Flash" at 310,76 size 148x16; Text 'A_Flash'
   Button "A_Bit" at 462,4 size 100x40; TextOff 'Text'
      Appearance <- "D_Bool"
   TextField "Label_A_Bit" at 462,76 size 148x16; Text 'A_Bit'
   Button "A_Bits" at 614,4 size 100x40; TextOff 'Text'
      Appearance <- "D_Bits"
   TextField "Label_A_Bits" at 614,76 size 148x16; Text 'A_Bits'
   Button "V_Range" at 6,96 size 100x40; TextOff 'Text'
      Visibility <- "D_Range"
   TextField "Label_V_Range" at 6,168 size 148x16; Text 'V_Range'
   Button "V_Bit" at 158,96 size 100x40; TextOff 'Text'
      Visibility <- "D_Vis"
   TextField "Label_V_Bit" at 158,168 size 148x16; Text 'V_Bit'
   Button "M_H" at 310,96 size 100x40; TextOff 'Text'
      HorizontalMovement <- "D_Pct"
   TextField "Label_M_H" at 310,168 size 148x16; Text 'M_H'
   Button "M_V" at 462,96 size 100x40; TextOff 'Text'
      VerticalMovement <- "D_Pct"
   TextField "Label_M_V" at 462,168 size 148x16; Text 'M_V'
   Button "M_D" at 614,96 size 100x40; TextOff 'Text'
      DiagonalMovement <- "D_Pct"
   TextField "Label_M_D" at 614,168 size 148x16; Text 'M_D'
   Button "M_Direct" at 6,188 size 100x40; TextOff 'Text'
      DirectMovement <- "D_X"
      DirectMovement <- "D_Y"
   TextField "Label_M_Direct" at 6,260 size 148x16; Text 'M_Direct'
   Button "E_Range" at 158,188 size 100x40; TextOff 'Text'
      ObjectEnable <- "D_Range"
   TextField "Label_E_Range" at 158,260 size 148x16; Text 'E_Range'
   Button "E_Bit" at 310,188 size 100x40; TextOff 'Text'
      ObjectEnable <- "D_En"
   TextField "Label_E_Bit" at 310,260 size 148x16; Text 'E_Bit'
   IOField "State" at 4,454 size 60x22; FormatPattern 9
      ProcessValue <- "D_State"
   Button "S1" at 70,454 size 40x22; TextOff 'S1'
      on Click: "SetS1"()
   Button "S2" at 114,454 size 40x22; TextOff 'S2'
      on Click: "SetS2"()
   Button "S3" at 158,454 size 40x22; TextOff 'S3'
      on Click: "SetS3"()
   Button "S4" at 202,454 size 40x22; TextOff 'S4'
      on Click: "SetS4"()
   Button "Next" at 756,454 size 40x22; TextOff 'Next'
      on Click: ActivateScreen("D_SymbolicIOField_1", 0)

screen "D_Circle_1" 800x480
   TextField "Label_Static" at 6,86 size 98x16; Text 'Static'
   Circle "A_Range" at 108,4 size 50x50
      Appearance <- "D_Range"
   TextField "Label_A_Range" at 108,86 size 98x16; Text 'A_Range'
   Circle "A_Flash" at 210,4 size 50x50
      Appearance <- "D_Range"
   TextField "Label_A_Flash" at 210,86 size 98x16; Text 'A_Flash'
   Circle "A_Bit" at 312,4 size 50x50
      Appearance <- "D_Bool"
   TextField "Label_A_Bit" at 312,86 size 98x16; Text 'A_Bit'
   Circle "A_Bits" at 414,4 size 50x50
      Appearance <- "D_Bits"
   TextField "Label_A_Bits" at 414,86 size 98x16; Text 'A_Bits'
   Circle "V_Range" at 516,4 size 50x50
      Visibility <- "D_Range"
   TextField "Label_V_Range" at 516,86 size 98x16; Text 'V_Range'
   Circle "V_Bit" at 618,4 size 50x50
      Visibility <- "D_Vis"
   TextField "Label_V_Bit" at 618,86 size 98x16; Text 'V_Bit'
   Circle "M_H" at 6,106 size 50x50
      HorizontalMovement <- "D_Pct"
   TextField "Label_M_H" at 6,188 size 98x16; Text 'M_H'
   Circle "M_V" at 108,106 size 50x50
      VerticalMovement <- "D_Pct"
   TextField "Label_M_V" at 108,188 size 98x16; Text 'M_V'
   Circle "M_D" at 210,106 size 50x50
      DiagonalMovement <- "D_Pct"
   TextField "Label_M_D" at 210,188 size 98x16; Text 'M_D'
   Circle "M_Direct" at 312,106 size 50x50
      DirectMovement <- "D_X"
      DirectMovement <- "D_Y"
   TextField "Label_M_Direct" at 312,188 size 98x16; Text 'M_Direct'
   Circle "E_Range" at 414,106 size 50x50
      ObjectEnable <- "D_Range"
   TextField "Label_E_Range" at 414,188 size 98x16; Text 'E_Range'
   Circle "E_Bit" at 516,106 size 50x50
      ObjectEnable <- "D_En"
   TextField "Label_E_Bit" at 516,188 size 98x16; Text 'E_Bit'
   IOField "State" at 4,454 size 60x22; FormatPattern 9
      ProcessValue <- "D_State"
   Button "S1" at 70,454 size 40x22; TextOff 'S1'
      on Click: "SetS1"()
   Button "S2" at 114,454 size 40x22; TextOff 'S2'
      on Click: "SetS2"()
   Button "S3" at 158,454 size 40x22; TextOff 'S3'
      on Click: "SetS3"()
   Button "S4" at 202,454 size 40x22; TextOff 'S4'
      on Click: "SetS4"()
   Button "Next" at 756,454 size 40x22; TextOff 'Next'
      on Click: ActivateScreen("D_Rectangle_1", 0)

screen "D_Clock_1" 800x480
   Clock "Static" at 6,4 size 150x150
   TextField "Label_Static" at 6,186 size 198x16; Text 'Static'
   Clock "A_Range" at 208,4 size 150x150
      Appearance <- "D_Range"
   TextField "Label_A_Range" at 208,186 size 198x16; Text 'A_Range'
   Clock "A_Flash" at 410,4 size 150x150
      Appearance <- "D_Range"
   TextField "Label_A_Flash" at 410,186 size 198x16; Text 'A_Flash'
   Clock "A_Bit" at 6,206 size 150x150
      Appearance <- "D_Bool"
   TextField "Label_A_Bit" at 6,388 size 198x16; Text 'A_Bit'
   Clock "A_Bits" at 208,206 size 150x150
      Appearance <- "D_Bits"
   TextField "Label_A_Bits" at 208,388 size 198x16; Text 'A_Bits'
   Clock "V_Range" at 410,206 size 150x150
      Visibility <- "D_Range"
   TextField "Label_V_Range" at 410,388 size 198x16; Text 'V_Range'
   IOField "State" at 4,454 size 60x22; FormatPattern 9
      ProcessValue <- "D_State"
   Button "S1" at 70,454 size 40x22; TextOff 'S1'
      on Click: "SetS1"()
   Button "S2" at 114,454 size 40x22; TextOff 'S2'
      on Click: "SetS2"()
   Button "S3" at 158,454 size 40x22; TextOff 'S3'
      on Click: "SetS3"()
   Button "S4" at 202,454 size 40x22; TextOff 'S4'
      on Click: "SetS4"()
   Button "Next" at 756,454 size 40x22; TextOff 'Next'
      on Click: ActivateScreen("D_Clock_2", 0)

screen "D_Clock_2" 800x480
   Clock "V_Bit" at 6,4 size 150x150
      Visibility <- "D_Vis"
   TextField "Label_V_Bit" at 6,186 size 198x16; Text 'V_Bit'
   Clock "M_H" at 208,4 size 150x150
      HorizontalMovement <- "D_Pct"
   TextField "Label_M_H" at 208,186 size 198x16; Text 'M_H'
   Clock "M_V" at 410,4 size 150x150
      VerticalMovement <- "D_Pct"
   TextField "Label_M_V" at 410,186 size 198x16; Text 'M_V'
   Clock "M_D" at 6,206 size 150x150
      DiagonalMovement <- "D_Pct"
   TextField "Label_M_D" at 6,388 size 198x16; Text 'M_D'
   Clock "M_Direct" at 208,206 size 150x150
      DirectMovement <- "D_X"
      DirectMovement <- "D_Y"
   TextField "Label_M_Direct" at 208,388 size 198x16; Text 'M_Direct'
   Clock "E_Range" at 410,206 size 150x150
      ObjectEnable <- "D_Range"
   TextField "Label_E_Range" at 410,388 size 198x16; Text 'E_Range'
   IOField "State" at 4,454 size 60x22; FormatPattern 9
      ProcessValue <- "D_State"
   Button "S1" at 70,454 size 40x22; TextOff 'S1'
      on Click: "SetS1"()
   Button "S2" at 114,454 size 40x22; TextOff 'S2'
      on Click: "SetS2"()
   Button "S3" at 158,454 size 40x22; TextOff 'S3'
      on Click: "SetS3"()
   Button "S4" at 202,454 size 40x22; TextOff 'S4'
      on Click: "SetS4"()
   Button "Next" at 756,454 size 40x22; TextOff 'Next'
      on Click: ActivateScreen("D_Clock_3", 0)

screen "D_Clock_3" 800x480
   Clock "E_Bit" at 6,4 size 150x150
      ObjectEnable <- "D_En"
   TextField "Label_E_Bit" at 6,186 size 198x16; Text 'E_Bit'
   IOField "State" at 4,454 size 60x22; FormatPattern 9
      ProcessValue <- "D_State"
   Button "S1" at 70,454 size 40x22; TextOff 'S1'
      on Click: "SetS1"()
   Button "S2" at 114,454 size 40x22; TextOff 'S2'
      on Click: "SetS2"()
   Button "S3" at 158,454 size 40x22; TextOff 'S3'
      on Click: "SetS3"()
   Button "S4" at 202,454 size 40x22; TextOff 'S4'
      on Click: "SetS4"()
   Button "Next" at 756,454 size 40x22; TextOff 'Next'
      on Click: ActivateScreen("D_Line_1", 0)

screen "D_DateTimeField_1" 800x480
   DateTimeField "Static" at 6,4 size 160x30
   TextField "Label_Static" at 6,66 size 208x16; Text 'Static'
   DateTimeField "A_Range" at 218,4 size 160x30
      Appearance <- "D_Range"
   TextField "Label_A_Range" at 218,66 size 208x16; Text 'A_Range'
   DateTimeField "A_Flash" at 430,4 size 160x30
      Appearance <- "D_Range"
   TextField "Label_A_Flash" at 430,66 size 208x16; Text 'A_Flash'
   DateTimeField "A_Bit" at 6,86 size 160x30
      Appearance <- "D_Bool"
   TextField "Label_A_Bit" at 6,148 size 208x16; Text 'A_Bit'
   DateTimeField "A_Bits" at 218,86 size 160x30
      Appearance <- "D_Bits"
   TextField "Label_A_Bits" at 218,148 size 208x16; Text 'A_Bits'
   DateTimeField "V_Range" at 430,86 size 160x30
      Visibility <- "D_Range"
   TextField "Label_V_Range" at 430,148 size 208x16; Text 'V_Range'
   DateTimeField "V_Bit" at 6,168 size 160x30
      Visibility <- "D_Vis"
   TextField "Label_V_Bit" at 6,230 size 208x16; Text 'V_Bit'
   DateTimeField "M_H" at 218,168 size 160x30
      HorizontalMovement <- "D_Pct"
   TextField "Label_M_H" at 218,230 size 208x16; Text 'M_H'
   DateTimeField "M_V" at 430,168 size 160x30
      VerticalMovement <- "D_Pct"
   TextField "Label_M_V" at 430,230 size 208x16; Text 'M_V'
   DateTimeField "M_D" at 6,250 size 160x30
      DiagonalMovement <- "D_Pct"
   TextField "Label_M_D" at 6,312 size 208x16; Text 'M_D'
   DateTimeField "M_Direct" at 218,250 size 160x30
      DirectMovement <- "D_X"
      DirectMovement <- "D_Y"
   TextField "Label_M_Direct" at 218,312 size 208x16; Text 'M_Direct'
   DateTimeField "E_Range" at 430,250 size 160x30
      ObjectEnable <- "D_Range"
   TextField "Label_E_Range" at 430,312 size 208x16; Text 'E_Range'
   DateTimeField "E_Bit" at 6,332 size 160x30
      ObjectEnable <- "D_En"
   TextField "Label_E_Bit" at 6,394 size 208x16; Text 'E_Bit'
   DateTimeField "PV_DateTime" at 218,332 size 160x30
      ProcessValue <- "D_DateTime"
   TextField "Label_PV_DateTime" at 218,394 size 208x16; Text 'PV_DateTime'
   IOField "State" at 4,454 size 60x22; FormatPattern 9
      ProcessValue <- "D_State"
   Button "S1" at 70,454 size 40x22; TextOff 'S1'
      on Click: "SetS1"()
   Button "S2" at 114,454 size 40x22; TextOff 'S2'
      on Click: "SetS2"()
   Button "S3" at 158,454 size 40x22; TextOff 'S3'
      on Click: "SetS3"()
   Button "S4" at 202,454 size 40x22; TextOff 'S4'
      on Click: "SetS4"()
   Button "Next" at 756,454 size 40x22; TextOff 'Next'
      on Click: ActivateScreen("D_Bar_1", 0)

screen "D_Ellipse_1" 800x480
   TextField "Label_Static" at 6,86 size 148x16; Text 'Static'
   Ellipse "A_Range" at 158,4 size 100x50
      Appearance <- "D_Range"
   TextField "Label_A_Range" at 158,86 size 148x16; Text 'A_Range'
   Ellipse "A_Flash" at 310,4 size 100x50
      Appearance <- "D_Range"
   TextField "Label_A_Flash" at 310,86 size 148x16; Text 'A_Flash'
   Ellipse "A_Bit" at 462,4 size 100x50
      Appearance <- "D_Bool"
   TextField "Label_A_Bit" at 462,86 size 148x16; Text 'A_Bit'
   Ellipse "A_Bits" at 614,4 size 100x50
      Appearance <- "D_Bits"
   TextField "Label_A_Bits" at 614,86 size 148x16; Text 'A_Bits'
   Ellipse "V_Range" at 6,106 size 100x50
      Visibility <- "D_Range"
   TextField "Label_V_Range" at 6,188 size 148x16; Text 'V_Range'
   Ellipse "V_Bit" at 158,106 size 100x50
      Visibility <- "D_Vis"
   TextField "Label_V_Bit" at 158,188 size 148x16; Text 'V_Bit'
   Ellipse "M_H" at 310,106 size 100x50
      HorizontalMovement <- "D_Pct"
   TextField "Label_M_H" at 310,188 size 148x16; Text 'M_H'
   Ellipse "M_V" at 462,106 size 100x50
      VerticalMovement <- "D_Pct"
   TextField "Label_M_V" at 462,188 size 148x16; Text 'M_V'
   Ellipse "M_D" at 614,106 size 100x50
      DiagonalMovement <- "D_Pct"
   TextField "Label_M_D" at 614,188 size 148x16; Text 'M_D'
   Ellipse "M_Direct" at 6,208 size 100x50
      DirectMovement <- "D_X"
      DirectMovement <- "D_Y"
   TextField "Label_M_Direct" at 6,290 size 148x16; Text 'M_Direct'
   Ellipse "E_Range" at 158,208 size 100x50
      ObjectEnable <- "D_Range"
   TextField "Label_E_Range" at 158,290 size 148x16; Text 'E_Range'
   Ellipse "E_Bit" at 310,208 size 100x50
      ObjectEnable <- "D_En"
   TextField "Label_E_Bit" at 310,290 size 148x16; Text 'E_Bit'
   IOField "State" at 4,454 size 60x22; FormatPattern 9
      ProcessValue <- "D_State"
   Button "S1" at 70,454 size 40x22; TextOff 'S1'
      on Click: "SetS1"()
   Button "S2" at 114,454 size 40x22; TextOff 'S2'
      on Click: "SetS2"()
   Button "S3" at 158,454 size 40x22; TextOff 'S3'
      on Click: "SetS3"()
   Button "S4" at 202,454 size 40x22; TextOff 'S4'
      on Click: "SetS4"()
   Button "Next" at 756,454 size 40x22; TextOff 'Next'
      on Click: ActivateScreen("D_Circle_1", 0)

screen "D_GraphicIOField_1" 800x480
   GraphicIOField "Static" at 6,4 size 60x60
   TextField "Label_Static" at 6,96 size 108x16; Text 'Static'
   GraphicIOField "A_Range" at 118,4 size 60x60
      Appearance <- "D_Range"
   TextField "Label_A_Range" at 118,96 size 108x16; Text 'A_Range'
   GraphicIOField "A_Flash" at 230,4 size 60x60
      Appearance <- "D_Range"
   TextField "Label_A_Flash" at 230,96 size 108x16; Text 'A_Flash'
   GraphicIOField "A_Bit" at 342,4 size 60x60
      Appearance <- "D_Bool"
   TextField "Label_A_Bit" at 342,96 size 108x16; Text 'A_Bit'
   GraphicIOField "A_Bits" at 454,4 size 60x60
      Appearance <- "D_Bits"
   TextField "Label_A_Bits" at 454,96 size 108x16; Text 'A_Bits'
   GraphicIOField "V_Range" at 566,4 size 60x60
      Visibility <- "D_Range"
   TextField "Label_V_Range" at 566,96 size 108x16; Text 'V_Range'
   GraphicIOField "V_Bit" at 678,4 size 60x60
      Visibility <- "D_Vis"
   TextField "Label_V_Bit" at 678,96 size 108x16; Text 'V_Bit'
   GraphicIOField "M_H" at 6,116 size 60x60
      HorizontalMovement <- "D_Pct"
   TextField "Label_M_H" at 6,208 size 108x16; Text 'M_H'
   GraphicIOField "M_V" at 118,116 size 60x60
      VerticalMovement <- "D_Pct"
   TextField "Label_M_V" at 118,208 size 108x16; Text 'M_V'
   GraphicIOField "M_D" at 230,116 size 60x60
      DiagonalMovement <- "D_Pct"
   TextField "Label_M_D" at 230,208 size 108x16; Text 'M_D'
   GraphicIOField "M_Direct" at 342,116 size 60x60
      DirectMovement <- "D_X"
      DirectMovement <- "D_Y"
   TextField "Label_M_Direct" at 342,208 size 108x16; Text 'M_Direct'
   GraphicIOField "E_Range" at 454,116 size 60x60
      ObjectEnable <- "D_Range"
   TextField "Label_E_Range" at 454,208 size 108x16; Text 'E_Range'
   GraphicIOField "E_Bit" at 566,116 size 60x60
      ObjectEnable <- "D_En"
   TextField "Label_E_Bit" at 566,208 size 108x16; Text 'E_Bit'
   IOField "State" at 4,454 size 60x22; FormatPattern 9
      ProcessValue <- "D_State"
   Button "S1" at 70,454 size 40x22; TextOff 'S1'
      on Click: "SetS1"()
   Button "S2" at 114,454 size 40x22; TextOff 'S2'
      on Click: "SetS2"()
   Button "S3" at 158,454 size 40x22; TextOff 'S3'
      on Click: "SetS3"()
   Button "S4" at 202,454 size 40x22; TextOff 'S4'
      on Click: "SetS4"()
   Button "Next" at 756,454 size 40x22; TextOff 'Next'
      on Click: ActivateScreen("D_DateTimeField_1", 0)

